(* IEC 61131-3 sources: daoli-st-library/DL_Algo (part 18) *)

(* ---- FB_DL_PidController.st ---- *)
(*==============================================================================
 * 组件名称 (Component)  : FB_DL_PidController
 * 所属子库 (Sublibrary) : DL_Algo
 * 当前版本 (Version)    : 1.0.1
 * 兼容性   (Platform)   : CODESYS 3.5 / TwinCAT 3 / 汇川 InoProShop / Machine Expert
 *                         仅依赖 Standard.library（R_TRIG），零厂商方言
 * 功能描述 (Function)   : 单回路通用离散 PID 控制器。位置式与增量式由独立布尔
 *                         bIncremental 选择（不堆模式枚举）；含控制死区、积分
 *                         分离（触限停积分）、两级抗积分饱和（条件积分 + 限幅
 *                         反算回填）、手自动无扰切换与跟踪回投。fKp 为负即反
 *                         作用（沿 OSCAT / 西门子惯例）。现场用途：温度 / 压力 /
 *                         流量单闭环调节主块，温控区与后续串级块的基石。
 * 开源溯源 (Origin)     : 原创实现。功能分类与参数域参考 OSCAT 基础库 FT_PIWL
 *                         反算抗饱和思想与西门子 CONT_C 公开语义描述，
 *                         未复制任何厂商源码，clean-room 重写。
 * 本文件内含       : TYPE  E_DL_PidState（配套枚举，归属 DL_Algo）
 *                    FB    FB_DL_PidController
 * 依赖     (Depends)    : 无 DL_ 内部依赖；Standard.library: R_TRIG
 * 红线自检 (Redline)    : R1 ✓ 零全局变量表与外部变量引用 ｜ R2 ✓ 零物理 IO 地址直写
 *                         R3 ✓ 纯 IEC 61131-3 ｜ R4 ✓ 防除零+钳位+非有限值防御
 *                         R5 ✓ 全变量中英双语同行注释 ｜ R6 ✓ 四态 ENUM+CASE+ELSE
 *                         R7 ✓ R_TRIG 实例主体最前部无条件刷新
 * 修订历史 (Revision)   :
 *   2026-11-15  v1.0.0  首版入库 · Round 04 · Level 1 DL_Algo
 *   2026-11-15  v1.0.1  阶段五终审精修：积分量纲统一为[%]；eIdle 补 bActive
 *                       清零；信息级码不置 bError；首扫与手自动历史同步防踢腿
 * 验收向量 (Acceptance) :
 *   V1 阶跃纯比例：fKp=2, tTi=T#0S, SP=50, PV=0 → fOut=rOutMax 触限
 *   V2 抗饱和：fKp=2, tTi=T#2S, SP=200 → 触上限后撤销阶跃，输出快速回落
 *      （积分已反算回填，无长时间停限）
 *   V3 无扰切换：手动 30.0 切自动首拍输出保持 30.0 连续
 *   V4 死区：fDeadband=5 且 |偏差|<5 → 输出保持不变
 *   V5 非有限值：fSetpoint 写入非法浮点 → 输出保持上一拍且 uErrorId=0002_0004
 *   V6 增量式：fKp=1, tTi=T#1S, 恒偏差 10 → fOut 单调爬升至上限后停
 *============================================================================*)
(*-----------------------------------------------------------------------------
 * 枚举: E_DL_PidState（归属 DL_Algo，与 FB_DL_PidController 同文件）
 * 含义: PID 控制器离散状态。数值步长留空位便于后续插态而不破坏已有工程。
 *----------------------------------------------------------------------------*)
TYPE E_DL_PidState :
(
    eIdle   := 0,    // 使能关：输出回输出下限，积分冻结 / Idle: enable off, output at low limit, integral frozen
    eAuto   := 10,   // 自动调节：闭环 PID 运算中 / Auto: closed-loop PID computation active
    eManual := 20,   // 手动模式：输出手动值，积分同步跟踪保证无扰 / Manual: output manual value, integral tracked for bumpless
    eFault  := 99    // 故障兜底态：非法状态进入，输出安全值 / Fault fallback: entered on illegal state, safe output
);
END_TYPE
(*==============================================================================
 * 功能块: FB_DL_PidController
 * 调用约定: 每个扫描周期无条件调用一次；bReset 上升沿清积分与故障。
 * 无状态泄漏: 全部状态驻留于实例私有 VAR，零全局引用，可多实例并行。
 * 工程披露: 微分项对偏差做一阶预滤波（滤波时间取 tTd 的 1/10），抑制微分尖峰。
 *============================================================================*)
FUNCTION_BLOCK FB_DL_PidController
VAR_INPUT
    bEnable      : BOOL := FALSE;     // 总使能，FALSE 时输出回输出下限 / Master enable, FALSE drives output to low limit
    bManual      : BOOL := FALSE;     // 手动模式选择，TRUE = 手动输出 / Manual mode select, TRUE = manual output
    fManualValue : REAL := 0.0;       // 手动输出值 [%]，越限自动钳位 / Manual output value [%], auto-clamped
    fSetpoint    : REAL := 0.0;       // 设定值 [EU] / Setpoint in engineering units
    fActual      : REAL := 0.0;       // 过程实际值 [EU] / Process actual value in engineering units
    fKp          : REAL := 1.0;       // 比例增益 [1]，负值 = 反作用 / Proportional gain, negative = reverse acting
    tTi          : TIME := T#2S;      // 积分时间 [s]，T#0S 表示纯 PD 无积分 / Integral time [s], T#0S = pure PD
    tTd          : TIME := T#0S;      // 微分时间 [s]，T#0S 关闭微分 / Derivative time [s], T#0S disables derivative
    fDeadband    : REAL := 0.0;       // 控制死区 [EU]，负值自动钳 0 / Control deadband [EU], negative clamped to 0
    bIncremental : BOOL := FALSE;     // TRUE = 增量式算法，FALSE = 位置式 / TRUE = incremental form, FALSE = positional
    rOutMin      : REAL := 0.0;       // 输出下限 [%] / Output lower limit in percent
    rOutMax      : REAL := 100.0;     // 输出上限 [%] / Output upper limit in percent
    tSampleTime  : TIME := T#100MS;   // 采样周期 [s]，小于 T#10MS 钳位 / Sample period, clamped to 10 ms minimum
    bTrack       : BOOL := FALSE;     // 跟踪使能，TRUE 时输出立即跟随跟踪值 / Track enable, output follows track value
    fTrackValue  : REAL := 0.0;       // 跟踪值 [%]，与输出同量纲，用于无扰投切 / Track value in percent, same unit as output
    bReset       : BOOL := FALSE;     // 复位信号，上升沿清积分与故障 / Reset, rising edge clears integral and fault
END_VAR
VAR_OUTPUT
    fOut         : REAL;              // 控制输出 [%] / Control output in percent
    fErr         : REAL;              // 偏差 = 设定 - 实际 [EU] / Error = setpoint minus actual
    fIntPart     : REAL;              // 积分分量 [%]，诊断用 / Integral component in percent, diagnostics
    bLimitHigh   : BOOL;              // 输出触上限标志 / Output saturated at upper limit flag
    bLimitLow    : BOOL;              // 输出触下限标志 / Output saturated at lower limit flag
    bActive      : BOOL;              // 自动调节进行中标志 / Auto regulation active flag
    bError       : BOOL;              // 故障标志，0 除外均置位 / Fault flag, set on any nonzero error code
    uErrorId     : UDINT;             // 故障码，0 = 无故障 / Error code, 0 = no error
END_VAR
VAR
    fErrPrev1    : REAL;              // 上一拍偏差（增量式历史） [EU] / Previous error for incremental form
    fErrPrev2    : REAL;              // 上上拍偏差（增量式历史） [EU] / Error two cycles ago for incremental form
    fErrF        : REAL;              // 微分预滤波后的偏差 [EU] / Prefiltered error for derivative term
    fErrFPrev    : REAL;              // 上一拍预滤波偏差 [EU] / Previous prefiltered error
    fbTrigReset  : R_TRIG;            // 复位信号上升沿检测实例 / Reset rising edge detector instance
    eState       : E_DL_PidState;     // 主状态机当前状态 / Current state of the main state machine
    bInit        : BOOL := TRUE;      // 历史同步标志，TRUE 触发历史同步（首扫即同步防踢腿）/ History sync flag, TRUE syncs histories on first scan
    fDt          : REAL;              // 生效采样周期 [s] / Effective sample period in seconds
    fLimLow      : REAL;              // 修复后的输出下限 [%] / Repaired output lower limit
    fLimHigh     : REAL;              // 修复后的输出上限 [%] / Repaired output upper limit
    fDeadbandEff : REAL;              // 钳位后的有效死区 [EU] / Clamped effective deadband
    fInt         : REAL;              // 积分累积 [%]，与输出同量纲 / Accumulated integral in percent, same unit as output
    fP           : REAL;              // 比例分量 [%] / Proportional component
    fD           : REAL;              // 微分分量 [%] / Derivative component
    fPre         : REAL;              // 抗饱和判定用预输出 [%] / Pre-output for anti-windup test
    fDelta       : REAL;              // 增量式单拍增量 [%] / Incremental delta of one cycle
    fTdS         : REAL;              // 微分时间换算秒 [s] / Derivative time in seconds
    fAlpha       : REAL;              // 微分预滤波权重 [0..1] / Derivative prefilter weight
    fManOut      : REAL;              // 钳位后的手动输出 [%] / Clamped manual output
    bSkipInt     : BOOL;              // 积分分离标志：触限且误差继续推进 / Conditional integration flag
END_VAR
VAR CONSTANT
    DL_PID_ERR_MAX : REAL := 1.0E10;  // 积分钳位上限 [%]，防浮点溢出的极端钳位 / Integral clamp ceiling [%], extreme guard against float overflow
END_VAR
(*------------------------------------------------------------------------------
 * 段 1｜无条件刷新区（红线 R7）：复位沿检测严禁进入任何 IF / CASE 分支
 *      Unconditional refresh zone (red line R7): edge detector outside IF / CASE
 *-----------------------------------------------------------------------------*)
fbTrigReset(CLK := bReset);
(*------------------------------------------------------------------------------
 * 段 2｜参数钳位与公共防御（不中断扫描，现场组态笔误不停机）
 *      Parameter clamping and common defenses, never stops the scan
 *-----------------------------------------------------------------------------*)
bError   := FALSE;                    // 每拍重算故障标志 / Recompute fault flag every cycle
uErrorId := 16#0002_0000;             // 每拍重算故障码 / Recompute error code every cycle
bLimitHigh := FALSE;                  // 触限标志每拍重算 / Saturation flags recomputed every cycle
bLimitLow  := FALSE;                  // 触限标志每拍重算 / Saturation flags recomputed every cycle
IF tSampleTime < T#10MS THEN
    fDt := 0.01;                      // 采样周期非法钳位为 0.01 s / Illegal sample period clamped to 0.01 s
    uErrorId := 16#0002_0002;         // 公共码：采样周期已钳位 / Common code: sample period clamped
ELSE
    fDt := TIME_TO_REAL(tSampleTime) / 1000.0;  // 采样周期换算为秒 [s] / Sample period converted to seconds
END_IF
IF rOutMin > rOutMax THEN
    fLimLow  := rOutMax;              // 上下限对调修复（下限取原上限） / Swapped limits after repair
    fLimHigh := rOutMin;              // 上下限对调修复（上限取原下限） / Swapped limits after repair
    uErrorId := 16#0002_0001;         // 公共码：参数越界已钳位 / Common code: parameter clamped
ELSE
    fLimLow  := rOutMin;              // 合法下限直通 / Valid lower limit passed through
    fLimHigh := rOutMax;              // 合法上限直通 / Valid upper limit passed through
END_IF
IF fDeadband < 0.0 THEN
    fDeadbandEff := 0.0;              // 死区负值钳 0 / Negative deadband clamped to zero
    uErrorId := 16#0002_0001;         // 公共码：参数越界已钳位 / Common code: parameter clamped
ELSE
    fDeadbandEff := fDeadband;        // 合法死区直通 / Valid deadband passed through
END_IF
(*------------------------------------------------------------------------------
 * 段 3｜复位处理：清积分、清增量式历史、清滤波偏差，故障归零
 *      Reset handling: clear integral, incremental history and filtered error
 *-----------------------------------------------------------------------------*)
IF fbTrigReset.Q THEN
    fInt       := 0.0;                // 清积分累积 [%] / Clear accumulated integral in percent
    fErrPrev1  := 0.0;                // 清上一拍偏差 / Clear previous error history
    fErrPrev2  := 0.0;                // 清上上拍偏差 / Clear two-cycle error history
    fErrF      := 0.0;                // 清滤波偏差 / Clear prefiltered error
    fErrFPrev  := 0.0;                // 清上拍滤波偏差 / Clear previous prefiltered error
    fOut       := fLimLow;            // 输出回安全下限 / Output to safe lower limit
    eState     := eIdle;              // 状态回空闲 / State back to idle
    bInit      := TRUE;               // 置首扫标志使下一拍同步历史 / Set init flag to resync history next cycle
END_IF
(*------------------------------------------------------------------------------
 * 段 4｜非有限值防御：设定值 / 过程值 / 手动值 / 跟踪值任一非法即拒绝本拍更新
 *      Non-finite defense: reject this cycle if any relevant input is invalid
 *-----------------------------------------------------------------------------*)
IF (fSetpoint <> fSetpoint) OR (ABS(fSetpoint) > 1.0E30)
   OR (fActual <> fActual) OR (ABS(fActual) > 1.0E30)
   OR (fManualValue <> fManualValue) OR (ABS(fManualValue) > 1.0E30)
   OR (fTrackValue <> fTrackValue) OR (ABS(fTrackValue) > 1.0E30) THEN
    bError   := TRUE;                 // 置故障标志 / Set fault flag
    uErrorId := 16#0002_0004;         // 公共码：输入非有限值已拒绝 / Common code: non-finite input rejected
    RETURN;                           // 保持上一拍输出与状态 / Hold previous output and state
END_IF
(*------------------------------------------------------------------------------
 * 段 5｜使能关断：输出回下限、积分冻结、状态回空闲（允许带电观察）
 *      Enable off: output to low limit, integral frozen, state back to idle
 *-----------------------------------------------------------------------------*)
IF NOT bEnable THEN
    eState  := eIdle;                 // 强制回空闲态 / Force idle state
    fOut    := fLimLow;               // 输出回下限安全值 / Output to safe low limit
    fErr    := fSetpoint - fActual;   // 偏差仍刷新供诊断 / Error still refreshed for diagnostics
    bActive := FALSE;                 // 调节未激活 / Regulation not active
    fIntPart:= fInt;                  // 保留积分分量供诊断 / Keep integral component for diagnostics
    RETURN;                           // 本拍结束 / End of this cycle
END_IF
(*------------------------------------------------------------------------------
 * 段 6｜主状态机（红线 R6）：ENUM + CASE + ELSE 兜底
 *      Main state machine: ENUM + CASE with mandatory ELSE fallback
 *-----------------------------------------------------------------------------*)
CASE eState OF
    eIdle:
        (* 空闲态：按手动 / 自动请求迁移，迁移前同步增量式历史防微分踢腿 *)
        (* Idle: migrate by mode request, sync incremental history before transfer *)
        bActive := FALSE;             // 空闲态激活标志清零防跨拍残留 / Clear active flag against stale carry-over
        fErr := fSetpoint - fActual;  // 计算原始偏差 [EU] / Raw error in engineering units
        IF ABS(fErr) < fDeadbandEff THEN
            fErr := 0.0;              // 死区内偏差按 0 处理 / Error inside deadband treated as zero
        END_IF
        IF bManual THEN
            eState := eManual;        // 请求手动 / Request manual mode
        ELSE
            eState := eAuto;          // 请求自动 / Request auto mode
        END_IF
    eAuto:
        (* 自动调节态：位置式或增量式 PID 闭环运算 + 两级抗饱和 *)
        (* Auto: positional or incremental closed-loop PID with two-stage anti-windup *)
        bActive := TRUE;              // 自动调节激活 / Auto regulation active
        fErr := fSetpoint - fActual;  // 原始偏差 [EU] / Raw error
        IF ABS(fErr) < fDeadbandEff THEN
            fErr := 0.0;              // 死区内偏差置 0 / Zero error inside deadband
        END_IF
        IF bInit THEN
            (* 首扫 / 复位后同步全部历史，杜绝上电尖峰与虚假微分 *)
            (* First scan / post-reset history sync, no power-up spike *)
            fErrF     := fErr;        // 滤波偏差同步 / Sync prefiltered error
            fErrFPrev := fErr;        // 上拍滤波偏差同步 / Sync previous prefiltered error
            fErrPrev1 := fErr;        // 增量式历史同步 / Sync incremental history
            fErrPrev2 := fErr;        // 增量式历史同步 / Sync incremental history
            bInit     := FALSE;       // 清首扫标志 / Clear first-scan flag
        END_IF
        fP := fKp * fErr;             // 比例项 [%] / Proportional term
        IF bTrack THEN
            (* 跟踪回投：输出立即跟随跟踪值，积分反算同步，恢复自动零扰动 *)
            (* Track mode: output follows track value, integral back-calculated in sync *)
            fOut    := LIMIT(fLimLow, fTrackValue, fLimHigh);   // 输出钳位跟随 / Clamped tracking output
            fInt    := fOut - fP - fD;                          // 积分反算同步 / Back-calculated integral
            fErrF   := fErr;        // 滤波偏差同步 / Sync prefiltered error
            fErrFPrev := fErr;      // 上拍滤波偏差同步 / Sync previous prefiltered error
            fErrPrev1 := fErr;      // 增量式历史同步 / Sync incremental history
            fErrPrev2 := fErr;      // 增量式历史同步 / Sync incremental history
            fIntPart := fInt;       // 诊断分量刷新 / Refresh diagnostic component
        ELSIF bIncremental THEN
            (* 增量式：PID 增量作用于输出累积，天然抗饱和由限幅兜底 *)
            (* Incremental form: PID delta applied to output accumulation *)
            fDelta := fKp * (fErr - fErrPrev1);                 // 比例增量 [%] / Proportional delta
            IF tTi > T#0S THEN
                fDelta := fDelta + fKp * fErr * fDt / (TIME_TO_REAL(tTi) / 1000.0);  // 积分增量 / Integral delta
            END_IF
            IF tTd > T#0S THEN
                fDelta := fDelta + fKp * (TIME_TO_REAL(tTd) / 1000.0) / fDt
                          * (fErr - 2.0 * fErrPrev1 + fErrPrev2);  // 微分增量 / Derivative delta
            END_IF
            fOut := LIMIT(fLimLow, fOut + fDelta, fLimHigh);    // 输出累积并限幅 / Accumulate and clamp
            fErrPrev2 := fErrPrev1;                             // 历史滚动 / Roll history
            fErrPrev1 := fErr;                                  // 历史滚动 / Roll history
            fIntPart  := fOut - fP - fD;                        // 诊断分量 / Diagnostic component
            IF ((fOut >= fLimHigh) AND (fDelta > 0.0))
               OR ((fOut <= fLimLow) AND (fDelta < 0.0)) THEN
                bLimitHigh := (fOut >= fLimHigh);               // 触上限标志 / Upper saturation flag
                bLimitLow  := (fOut <= fLimLow);                // 触下限标志 / Lower saturation flag
                IF uErrorId = 16#0002_0000 THEN
                    uErrorId := 16#0002_0101;                   // 信息级：输出饱和提示 / Info: output saturated
                END_IF
            END_IF
        ELSE
            (* 位置式：先做微分预滤波，再做积分分离与两级抗饱和 *)
            (* Positional: derivative prefilter, then conditional integration and back-calc *)
            IF tTd > T#0S THEN
                fTdS   := TIME_TO_REAL(tTd) / 1000.0;           // 微分时间换算秒 [s] / Derivative time in seconds
                fAlpha := fDt / (0.1 * fTdS + fDt);             // 预滤波权重 [0..1] / Prefilter weight
                fErrF  := fErrF + fAlpha * (fErr - fErrF);      // 一阶预滤波递推 / First-order prefilter recursion
                fD     := fKp * fTdS / fDt * (fErrF - fErrFPrev);  // 微分项 [%] / Derivative term
                fErrFPrev := fErrF;                             // 滚动滤波历史 / Roll filtered history
            ELSE
                fD        := 0.0;                               // 微分关闭 / Derivative disabled
                fErrF     := fErr;                              // 滤波偏差直通 / Prefiltered error follows
                fErrFPrev := fErr;                              // 上拍滤波偏差同步 / Sync previous value
            END_IF
            fPre := fP + fD + fInt;                             // 当前积分下的预输出 [%] / Pre-output with current integral
            bSkipInt := (fPre > fLimHigh AND fErr > 0.0)
                     OR (fPre < fLimLow  AND fErr < 0.0);       // 积分分离判定 / Conditional integration test
            IF (tTi > T#0S) AND (NOT bSkipInt) THEN
                fInt := fInt + fKp * fErr * fDt / (TIME_TO_REAL(tTi) / 1000.0);  // 条件积分 / Conditional integration
            END_IF
            fInt := LIMIT(-DL_PID_ERR_MAX, fInt, DL_PID_ERR_MAX);  // 积分钳位防溢出 / Clamp integral against overflow
            fPre := fP + fD + fInt;                             // 二次合成预输出 [%] / Recomposed pre-output
            IF fPre > fLimHigh THEN
                fOut := fLimHigh;                               // 输出钳上限 / Output at upper limit
                fInt := fLimHigh - fP - fD;                     // 反算回填积分 / Back-calculated integral
                bLimitHigh := TRUE;                             // 触上限标志 / Upper saturation flag
                IF uErrorId = 16#0002_0000 THEN
                    uErrorId := 16#0002_0101;                   // 信息级：输出饱和提示 / Info: output saturated
                END_IF
            ELSIF fPre < fLimLow THEN
                fOut := fLimLow;                                // 输出钳下限 / Output at lower limit
                fInt := fLimLow - fP - fD;                      // 反算回填积分 / Back-calculated integral
                bLimitLow := TRUE;                              // 触下限标志 / Lower saturation flag
                IF uErrorId = 16#0002_0000 THEN
                    uErrorId := 16#0002_0101;                   // 信息级：输出饱和提示 / Info: output saturated
                END_IF
            ELSE
                fOut := fPre;                                   // 正常输出 / Normal output
            END_IF
            fIntPart := fInt;                                   // 诊断分量刷新 / Refresh diagnostic component
        END_IF
        IF bManual THEN
            eState := eManual;                                  // 切手动 / Switch to manual
        END_IF
    eManual:
        (* 手动态：输出手动值（钳位），积分反算同步保证回自动瞬间输出连续 *)
        (* Manual: clamped manual output, integral back-calculated for bumpless return *)
        bActive := FALSE;                                       // 自动调节未激活 / Auto not active
        fErr := fSetpoint - fActual;                            // 偏差仍计算供诊断 / Error for diagnostics
        IF ABS(fErr) < fDeadbandEff THEN
            fErr := 0.0;                                        // 死区内偏差置 0 / Zero inside deadband
        END_IF
        (* 手动期间持续同步微分与增量式历史，杜绝切回自动瞬间的踢腿 *)
        (* Keep syncing derivative and incremental history in manual, no kick on auto return *)
        fErrF     := fErr;                                      // 微分滤波偏差同步 / Sync prefiltered error
        fErrFPrev := fErr;                                      // 上拍滤波偏差同步 / Sync previous prefiltered error
        fErrPrev1 := fErr;                                      // 增量式历史同步 / Sync incremental history
        fErrPrev2 := fErr;                                      // 增量式历史同步 / Sync incremental history
        fP := fKp * fErr;                                       // 比例项 [%] / Proportional term
        fD := 0.0;                                              // 手动下微分置 0 / Derivative zero in manual
        fManOut := LIMIT(fLimLow, fManualValue, fLimHigh);      // 手动值钳位 / Clamped manual value
        IF fManualValue > fLimHigh OR fManualValue < fLimLow THEN
            IF uErrorId = 16#0002_0000 THEN
                uErrorId := 16#0002_0102;                       // 手动值超限已钳位 / Manual value clamped
            END_IF
        END_IF
        fOut      := fManOut;                                   // 输出手动值 / Output manual value
        fInt      := fManOut - fP - fD;                         // 积分反算同步 / Back-calculated integral
        fInt      := LIMIT(-DL_PID_ERR_MAX, fInt, DL_PID_ERR_MAX);  // 积分钳位 / Clamp integral
        fIntPart  := fInt;                                      // 诊断分量刷新 / Refresh diagnostic component
        IF bTrack THEN
            fOut := LIMIT(fLimLow, fTrackValue, fLimHigh);      // 跟踪值优先 / Track value takes priority
            fInt := fOut - fP - fD;                             // 积分同步 / Integral in sync
        END_IF
        IF bInit THEN
            fErrF     := fErr;                                  // 滤波偏差同步 / Sync prefiltered error
            fErrFPrev := fErr;                                  // 上拍滤波偏差同步 / Sync previous value
            fErrPrev1 := fErr;                                  // 增量式历史同步 / Sync history
            fErrPrev2 := fErr;                                  // 增量式历史同步 / Sync history
            bInit     := FALSE;                                 // 清首扫标志 / Clear first-scan flag
        END_IF
        IF NOT bManual THEN
            eState := eAuto;                                    // 切自动 / Switch to auto
        END_IF
    eFault:
        (* 故障兜底态：输出安全下限，等待复位沿解除 *)
        (* Fault fallback: safe low-limit output, released by reset edge *)
        fOut    := fLimLow;                                     // 安全输出 / Safe output
        bActive := FALSE;                                       // 调节未激活 / Not active
    ELSE
        (* 非法状态拦截：任何未定义状态一律进故障兜底，不做隐式恢复 *)
        (* Illegal state interception: any undefined state goes to fault fallback *)
        eState   := eFault;                                     // 进故障态 / Enter fault state
        bError   := TRUE;                                       // 置故障标志 / Set fault flag
        uErrorId := 16#0002_0005;                               // 非法状态兜底码 / Illegal state fallback code
        fOut     := fLimLow;                                    // 安全输出 / Safe output
END_CASE;
(* 信息级码（0101 输出饱和 / 0102 手动值钳位）不置故障标志，防下游报警误动作 *)
(* Info-level codes (saturation / manual clamp) never raise the fault flag *)
bError := (uErrorId <> 16#0002_0000) AND (uErrorId <> 16#0002_0101)
          AND (uErrorId <> 16#0002_0102);                        // 非信息级码才置故障 / Fault flag only on non-info codes
END_FUNCTION_BLOCK

(* ---- FB_DL_PidGainScheduler.st ---- *)
(*==============================================================================
 * 组件名称 (Component)  : FB_DL_PidGainScheduler
 * 溯源说明 (Provenance) : 道莅 clean-room 防御性实现（LGF Technology 深化 + 规划新增线）
 * 所属子库 (Sublibrary) : DL_Algo / ControlParams
 * 当前版本 (Version)    : 1.0.0
 * 兼容性   (Platform)   : CODESYS 3.5 / TwinCAT 3 / 汇川 InoProShop；
 *                         纯 IEC 61131-3（第 3 版），零标准库依赖
 * 组件分类 (Category)   : 功能块（FUNCTION_BLOCK）· 增益调度查表插值
 * 功能一句话 (Summary)  : 按调度变量查增益表线性插值输出 Kp/Ti/Td，仅出参数不控回路。
 * 边界与安全 (Boundary) : ①调度变量低于首点/高于末点 → 端点钳位并置码 3705；
 *                         ②表未按 fVar 严格升序 → 码 3701 且 bHoldLast 生效保持上次输出；
 *                         ③调度变量 NaN → 码 3702 保持上次输出；
 *                         ④表点数不足 2 → 视同表非法（3701 复用）；
 *                         ⑤本件只产出参数，不内嵌控制回路（与 PID 件正交解耦）。
 * 错误码    : 16#0002_3701 增益表非法（未升序或点数不足）——故障级（持续态）
 *             16#0002_3702 调度变量 NaN（保持上次输出）——故障级（持续态）
 *             16#0002_3705 端点钳位发生——信息级（持续态）
 * 码位总账  : 16#0002_3701 用 / 16#0002_3702 用 / 16#0002_3705 用
 * 修改记录  : v1.0.0 R26 初版
 *==============================================================================*)
TYPE ST_DL_GainPoint :
STRUCT
    fVar : LREAL; // 调度变量锚点 / Scheduling variable anchor
    fKp  : LREAL; // 该锚点比例增益 / Proportional gain at anchor
    fTi  : LREAL; // 该锚点积分时间 [s] / Integral time at anchor [s]
    fTd  : LREAL; // 该锚点微分时间 [s] / Derivative time at anchor [s]
END_STRUCT
END_TYPE

FUNCTION_BLOCK FB_DL_PidGainScheduler
VAR_INPUT
    fSchedVar  : LREAL; // 调度变量（如流量/温度工况）/ Scheduling variable
    bEnable    : BOOL;  // 使能：FALSE 保持上次输出 / Enable: FALSE holds last output
    bHoldLast  : BOOL;  // 表非法时保持上次输出 / Hold last output on illegal table
END_VAR
VAR_IN_OUT
    aGainTable : ARRAY[*] OF ST_DL_GainPoint; // 增益表，须按 fVar 升序 / Gain table, ascending by fVar
END_VAR
VAR_OUTPUT
    fKp   : LREAL; // 插值输出比例增益 / Interpolated proportional gain
    fTi   : LREAL; // 插值输出积分时间 [s] / Interpolated integral time [s]
    fTd   : LREAL; // 插值输出微分时间 [s] / Interpolated derivative time [s]
    eErr  : UDINT; // 本周期错误码，0=无错 / Error code this cycle, 0 = none
END_VAR
VAR
    nPts    : INT;  // 表点数 / Table point count
    i       : INT;  // 分段搜索游标 / Segment search cursor
    fDen    : LREAL; // 分段分母（前判零）/ Segment denominator (zero-guarded)
    fRatio  : LREAL; // 段内插值比例 / Interpolation ratio
    bTableOk: BOOL; // 表合法性中间判据 / Table legality intermediate
    bHold   : BOOL; // 本拍保持输出判据 / Hold-output predicate this cycle
END_VAR

// ---------- 周期起点：错误码清零（持续态随后重置） ----------
eErr := 0;
bHold := FALSE;

// ---------- 使能为假：纯保持，不查表不刷新 ----------
IF NOT bEnable THEN
    bHold := TRUE;                            // 保持上次输出 / Hold last output
ELSE
    // ---------- 表点数与单调性防御 ----------
    nPts := UPPER_BOUND(aGainTable, 1) + 1;   // 表点数 / Point count
    bTableOk := nPts >= 2;                    // 至少两点 / At least two points
    IF bTableOk THEN
        FOR i := 0 TO nPts - 2 DO
            IF NOT (aGainTable[i].fVar < aGainTable[i + 1].fVar) THEN
                bTableOk := FALSE;            // 严格升序被破坏 / Strict order violated
            END_IF
        END_FOR
    END_IF
    IF NOT bTableOk THEN
        eErr  := 16#0002_3701;                // 表非法码 / Illegal table code
        bHold := bHoldLast;                   // 按调用方策略保持 / Hold per caller policy
    ELSE
        // ---------- NaN 调度变量：保持 ----------
        IF fSchedVar <> fSchedVar THEN
            eErr  := 16#0002_3702;            // NaN 码 / NaN code
            bHold := TRUE;                    // 强制保持 / Forced hold
        ELSE
            // ---------- 端点钳位与段内插值 ----------
            IF fSchedVar <= aGainTable[0].fVar THEN
                fKp := aGainTable[0].fKp;     // 低于首点钳端点 / Below first: clamp endpoint
                fTi := aGainTable[0].fTi;
                fTd := aGainTable[0].fTd;
                IF fSchedVar < aGainTable[0].fVar THEN
                    eErr := 16#0002_3705;     // 端点钳位码 / Endpoint clamp code
                END_IF
            ELSIF fSchedVar >= aGainTable[nPts - 1].fVar THEN
                fKp := aGainTable[nPts - 1].fKp; // 高于末点钳端点 / Above last: clamp endpoint
                fTi := aGainTable[nPts - 1].fTi;
                fTd := aGainTable[nPts - 1].fTd;
                IF fSchedVar > aGainTable[nPts - 1].fVar THEN
                    eErr := 16#0002_3705;     // 端点钳位码 / Endpoint clamp code
                END_IF
            ELSE
                i := 0;
                WHILE (i < nPts - 2) AND (fSchedVar > aGainTable[i + 1].fVar) DO
                    i := i + 1;               // 定位所在段 / Locate segment
                END_WHILE
                fDen := aGainTable[i + 1].fVar - aGainTable[i].fVar; // 段宽 / Segment width
                IF fDen > 0.0 THEN
                    fRatio := (fSchedVar - aGainTable[i].fVar) / fDen; // 除法前判零 / Zero-guarded divide
                    fKp := aGainTable[i].fKp + fRatio * (aGainTable[i + 1].fKp - aGainTable[i].fKp);
                    fTi := aGainTable[i].fTi + fRatio * (aGainTable[i + 1].fTi - aGainTable[i].fTi);
                    fTd := aGainTable[i].fTd + fRatio * (aGainTable[i + 1].fTd - aGainTable[i].fTd);
                ELSE
                    fKp := aGainTable[i].fKp; // 段宽为零防御取左点 / Zero-width defensive left point
                    fTi := aGainTable[i].fTi;
                    fTd := aGainTable[i].fTd;
                END_IF
            END_IF
        END_IF
    END_IF
END_IF

// ---------- 保持路径显式化：bHold 时三输出不动（锁存语义注释） ----------
// bHold=TRUE 期间 fKp/fTi/fTd 为上次有效锁存值，内部不引入实时镜像副本，
// 输出与内部判定共用同一组锁存变量，避免双口径混用。

END_FUNCTION_BLOCK

(* ---- FB_DL_PidParamDriftAudit.st ---- *)
(*
  Name        : FB_DL_PidParamDriftAudit
  Category    : DL_Algo
  Version     : 1.0.1
  Purpose     : 整定参数漂移审计：逐拍比对现行 Kp/Ti/Td 与基准快照，按相对容差判漂移并累计越差次数，供「谁改了参数」留痕；/ Audit PID parameter drift: compare live Kp/Ti/Td against baseline snapshots with relative tolerance, accumulate excursions for an auditable trail
  溯源        : 借 t2-3-风格指南·审计 的分类/参数域组织，clean-room 实现
  Boundary    : ① 基准近零分支：|基准| <= eps 时相对偏差无定义，改走绝对差判据（fTolAbs），不产生除零/Inf；
                ② 现行与基准同为近零 → 判无漂移（0/0 语义按「一致」处理）；
                ③ 容差与近零判据全部 ABS 差比较，禁 `=`/`<>`；
                ④ 越差计数饱和累加，防 UDINT 回绕；
                ⑤ 本件只审计不改参数，输出仅供上位留痕（属主边界）。
  修订记录    : 2026-11-20 v1.0.1：六参数有限性闸补 Inf 差判（NaN+Inf 双闸，R52-05）；bDriftAny 改由三确认位 OR 同源重算（R52-06）；_fHun 迁入 VAR CONSTANT c_fHun 收口魔法数。
*)
TYPE E_DL_PdaState :
(
    eIdle  := 0,                             (* 未使能 / Disabled *)
    eAudit := 10,                            (* 审计运行 / Auditing *)
    eFault := 90                             (* 故障锁存相 / Fault latched *)
);
END_TYPE

TYPE E_DL_PdaCause :
(
    eNone       := 0,                        (* 无故障成因 / No cause *)
    eCfgIllegal := 1,                        (* 组态非法：容差/参考值越域 / Illegal config *)
    ePhaseBad   := 2                         (* 非法相位兜底 / Illegal phase fallback *)
);
END_TYPE

FUNCTION_BLOCK FB_DL_PidParamDriftAudit
VAR_INPUT
    fKp        : REAL := 1.0;                (* 现行比例增益 [-] / Live proportional gain *)
    fTi        : REAL := 1.0;                (* 现行积分时间，P 模式可为 0 [s] / Live integral time, 0 allowed *)
    fTd        : REAL := 0.0;                (* 现行微分时间，P/PI 模式可为 0 [s] / Live derivative time, 0 allowed *)
    fKpRef     : REAL := 1.0;                (* 基准比例增益（签核快照）[-] / Baseline proportional gain *)
    fTiRef     : REAL := 1.0;                (* 基准积分时间 [s] / Baseline integral time *)
    fTdRef     : REAL := 0.0;                (* 基准微分时间 [s] / Baseline derivative time *)
    fTolRel    : REAL := 0.05;               (* 相对漂移容差（5% = 0.05），域 > 0 [-] / Relative tolerance, > 0 *)
    fTolAbs    : REAL := 0.01;               (* 基准近零时改用的绝对差容差，域 > 0 [参数单位] / Absolute tolerance for near-zero baselines *)
    nConfirm   : INT := 3;                   (* 越差确认拍数，域 >= 1 [拍] / Consecutive excursion scans to confirm *)
    bEnable    : BOOL := TRUE;               (* 审计使能 [-] / Enable *)
    bReset      : BOOL := FALSE;             (* 复位命令，上升沿清漂移标志与计数 [-] / Reset command *)
END_VAR
VAR_OUTPUT
    fDriftKp   : REAL;                       (* Kp 相对漂移（% / 近零基准时为绝对差）[%] / Kp drift *)
    fDriftTi   : REAL;                       (* Ti 相对漂移 [%] / Ti drift *)
    fDriftTd   : REAL;                       (* Td 相对漂移 [%] / Td drift *)
    bDriftKp   : BOOL;                       (* Kp 越差确认位 [-] / Kp drift confirmed *)
    bDriftTi   : BOOL;                       (* Ti 越差确认位 [-] / Ti drift confirmed *)
    bDriftTd   : BOOL;                       (* Td 越差确认位 [-] / Td drift confirmed *)
    bDriftAny  : BOOL;                       (* 任一参数越差（汇总位）[-] / Any parameter drifted *)
    nDriftCnt  : UDINT;                      (* 累计确认越差次数（饱和）[-] / Confirmed drift count, saturated *)
    eState     : E_DL_PdaState;              (* 状态出口 / State outlet *)
    eCause     : E_DL_PdaCause;              (* 故障成因出口（R190 归因唯一） / Fault cause outlet *)
    bError     : BOOL;                       (* 故障锁存标志 [-] / Fault latch flag *)
END_VAR
VAR
    _eState  : E_DL_PdaState := E_DL_PdaState.eIdle;     (* 内部相位（CASE 唯一写入目标） / Internal phase *)
    _eCause  : E_DL_PdaCause := E_DL_PdaCause.eNone;     (* 故障成因锁存量 / Latched cause *)
    rtReset  : R_TRIG;                       (* 复位沿实例，段 0 无条件调用 / Reset edge instance *)
    _bFault  : BOOL;                         (* 故障锁存位 / Latched fault bit *)
    _bCfgBad : BOOL;                         (* 组态非法当拍量 / Illegal config this scan *)
    _bFinite : BOOL;                         (* 六参数有限性联合闸 / Finiteness of all six parameters *)
    _bExKp   : BOOL;                         (* Kp 当拍越差（未确认） / Kp excursion this scan *)
    _bExTi   : BOOL;                         (* Ti 当拍越差 / Ti excursion this scan *)
    _bExTd   : BOOL;                         (* Td 当拍越差 / Td excursion this scan *)
    _bAny    : BOOL;                         (* 任一当拍越差 / Any excursion this scan *)
    _nHold   : INT;                          (* 越差连续拍计数 [-] / Consecutive excursion counter *)
    _fDkp    : REAL;                         (* Kp 偏差绝对值/相对值中间量 [%] / Kp deviation intermediate *)
    _fDti    : REAL;                         (* Ti 偏差中间量 [%] / Ti deviation intermediate *)
    _fDtd    : REAL;                         (* Td 偏差中间量 [%] / Td deviation intermediate *)
END_VAR
VAR CONSTANT
    DL_PDA_EPS    : REAL  := 1.0E-6;         (* 近零/容差判零容差（REAL 量级）[-] / Epsilon *)
    DL_PDA_CNTMAX : UDINT := 4294967295;     (* 计数饱和上限（R28）[-] / Count saturation cap *)
    DL_PDA_NMAX   : INT   := 100;            (* 确认拍数上限（防长时间不判）[拍] / Confirm scans cap *)
    c_fHun        : LREAL := 100.0;          (* 百分数换算常量（v1.0.1 由 VAR 迁入收口）[-] / Percent scale constant *)
END_VAR

(* —— 段 0：当拍判据派生 + 实例无条件刷新（R228A） —— *)
_bCfgBad := (fTolRel <= DL_PDA_EPS) OR (fTolAbs <= DL_PDA_EPS)                 (* 容差正域闸（两口径均须有效） / Tolerance gates *)
            OR (nConfirm < 1) OR (nConfirm > DL_PDA_NMAX);                     (* 确认拍数域闸 / Confirm-count gate *)
rtReset(CLK := bReset);                                                        (* 复位沿每拍必调 / Reset edge every scan *)
_bFinite := (fKp = fKp) AND ((fKp - fKp) = (fKp - fKp))                        (* Kp NaN 自反 + Inf 差判闸（v1.0.1）/ Kp NaN and Inf gates *)
            AND (fTi = fTi) AND ((fTi - fTi) = (fTi - fTi))                    (* Ti NaN 自反 + Inf 差判闸 / Ti NaN and Inf gates *)
            AND (fTd = fTd) AND ((fTd - fTd) = (fTd - fTd))                    (* Td NaN 自反 + Inf 差判闸 / Td NaN and Inf gates *)
            AND (fKpRef = fKpRef) AND ((fKpRef - fKpRef) = (fKpRef - fKpRef))  (* 基准 Kp NaN + Inf 闸 / Baseline Kp NaN and Inf gates *)
            AND (fTiRef = fTiRef) AND ((fTiRef - fTiRef) = (fTiRef - fTiRef))  (* 基准 Ti NaN + Inf 闸 / Baseline Ti NaN and Inf gates *)
            AND (fTdRef = fTdRef) AND ((fTdRef - fTdRef) = (fTdRef - fTdRef)); (* 基准 Td NaN + Inf 闸（Inf-Inf→NaN 漏报收口）/ Baseline Td NaN and Inf gates *)

(* —— 段 1：单拍量预清零（R107） —— *)
_bExKp := FALSE;                                                               (* Kp 越差预清 / Kp excursion preset *)
_bExTi := FALSE;                                                               (* Ti 越差预清 / Ti excursion preset *)
_bExTd := FALSE;                                                               (* Td 越差预清 / Td excursion preset *)
_bAny := FALSE;                                                                (* 汇总位预清 / Any preset *)
(* bDriftAny 不再每拍独立预清：改由段 5 由三确认位 OR 同源重算（v1.0.1，R52-06 汇总不回落） *)

(* —— 段 2：复位沿处理（作用域：清故障 + 清三个确认位 + 清计数 + 迁 eIdle，R283 逐项声明） —— *)
IF rtReset.Q THEN
    _bFault := FALSE;                                                          (* 清故障锁存 / Clear fault *)
    _eCause := E_DL_PdaCause.eNone;                                            (* 清成因 / Clear cause *)
    bDriftKp := FALSE;                                                         (* 清 Kp 确认位 / Clear Kp confirm *)
    bDriftTi := FALSE;                                                         (* 清 Ti 确认位 / Clear Ti confirm *)
    bDriftTd := FALSE;                                                         (* 清 Td 确认位 / Clear Td confirm *)
    nDriftCnt := 0;                                                            (* 清越差计数 / Clear count *)
    _nHold := 0;                                                               (* 清连续拍计数 / Clear hold counter *)
    fDriftKp := 0.0;                                                           (* 清 Kp 漂移出口 / Clear Kp drift outlet *)
    fDriftTi := 0.0;                                                           (* 清 Ti 漂移出口 / Clear Ti drift outlet *)
    fDriftTd := 0.0;                                                           (* 清 Td 漂移出口 / Clear Td drift outlet *)
    _eState := E_DL_PdaState.eIdle;                                            (* 迁未使能相 / Back to idle *)
END_IF

(* —— 段 3：组态故障锁存（锁存至复位沿，R189） —— *)
IF _bCfgBad AND NOT _bFault THEN
    _bFault := TRUE;                                                           (* 锁存故障位 / Latch fault *)
    _eCause := E_DL_PdaCause.eCfgIllegal;                                      (* 成因：组态非法 / Cause: illegal config *)
    _eState := E_DL_PdaState.eFault;                                           (* 同步迁故障相 / Migrate to fault *)
END_IF

(* —— 段 4：CASE 主状态机（ELSE 兜底迁 eFault，红线 6） —— *)
CASE _eState OF
    E_DL_PdaState.eIdle:                                                       (* 未使能：不审计，出口保持 / Disabled *)
        _nHold := 0;                                                           (* 失能清连续计数（防隐性回夹） / Clear hold *)
        IF bEnable AND NOT _bFault THEN
            _eState := E_DL_PdaState.eAudit;                                   (* 使能进入审计 / Enter audit *)
        END_IF
    E_DL_PdaState.eAudit:                                                      (* 审计相：三参数双口径比对 / Auditing *)
        IF NOT bEnable THEN
            _eState := E_DL_PdaState.eIdle;                                    (* 失能回未使能 / Back to idle *)
        ELSIF _bFinite THEN
            IF ABS(fKpRef) > DL_PDA_EPS THEN
                _fDkp := LREAL_TO_REAL(ABS(fKp - fKpRef) / ABS(fKpRef) * c_fHun);   (* 相对漂移 %：除子已过闸，显式窄化转换 / Relative drift, divisor gated *)
                _bExKp := _fDkp > LREAL_TO_REAL(fTolRel * c_fHun);             (* 越差判据：相对口径 / Excursion, relative *)
            ELSE
                _fDkp := ABS(fKp - fKpRef);                                    (* 基准近零：退化为绝对差（边界①） / Near-zero baseline: absolute *)
                _bExKp := _fDkp > fTolAbs;                                     (* 越差判据：绝对口径 / Excursion, absolute *)
            END_IF
            IF ABS(fTiRef) > DL_PDA_EPS THEN
                _fDti := LREAL_TO_REAL(ABS(fTi - fTiRef) / ABS(fTiRef) * c_fHun);   (* Ti 相对漂移 % / Ti relative drift *)
                _bExTi := _fDti > LREAL_TO_REAL(fTolRel * c_fHun);             (* Ti 越差判据 / Ti excursion *)
            ELSE
                _fDti := ABS(fTi - fTiRef);                                    (* Ti 基准为 0：绝对差（P 模式常见） / Ti near-zero: absolute *)
                _bExTi := _fDti > fTolAbs;                                     (* Ti 越差判据（绝对） / Ti excursion, absolute *)
            END_IF
            IF ABS(fTdRef) > DL_PDA_EPS THEN
                _fDtd := LREAL_TO_REAL(ABS(fTd - fTdRef) / ABS(fTdRef) * c_fHun);   (* Td 相对漂移 % / Td relative drift *)
                _bExTd := _fDtd > LREAL_TO_REAL(fTolRel * c_fHun);             (* Td 越差判据 / Td excursion *)
            ELSE
                _fDtd := ABS(fTd - fTdRef);                                    (* Td 基准为 0：绝对差 / Td near-zero: absolute *)
                _bExTd := _fDtd > fTolAbs;                                     (* Td 越差判据（绝对） / Td excursion, absolute *)
            END_IF
            fDriftKp := _fDkp;                                                 (* Kp 漂移出口（实时派生） / Kp drift outlet *)
            fDriftTi := _fDti;                                                 (* Ti 漂移出口 / Ti drift outlet *)
            fDriftTd := _fDtd;                                                 (* Td 漂移出口 / Td drift outlet *)
            _bAny := _bExKp OR _bExTi OR _bExTd;                               (* 任一越差汇总 / Any excursion *)
            IF _bAny THEN
                _nHold := _nHold + 1;                                          (* 连续越差拍递增 / Increment hold *)
            ELSE
                _nHold := 0;                                                   (* 有拍未越差即清零（降抖） / Reset on clean scan *)
            END_IF
            IF _nHold >= nConfirm THEN                                         (* 连续确认拍数到齐 / Confirm reached *)
                IF _bExKp THEN
                    bDriftKp := TRUE;                                          (* Kp 确认位锁存 / Latch Kp confirm *)
                END_IF
                IF _bExTi THEN
                    bDriftTi := TRUE;                                          (* Ti 确认位锁存 / Latch Ti confirm *)
                END_IF
                IF _bExTd THEN
                    bDriftTd := TRUE;                                          (* Td 确认位锁存 / Latch Td confirm *)
                END_IF
                IF nDriftCnt < DL_PDA_CNTMAX THEN
                    nDriftCnt := nDriftCnt + 1;                                (* 越差事件净额 +1（同拍多次不叠加） / Net +1 per confirmed event *)
                END_IF
                _nHold := 0;                                                   (* 计数归零，下一轮重新累积 / Restart accumulation *)
            END_IF
        END_IF                                                                 (* 非有限参数：本拍不判（保留确认位） / Non-finite: skip verdict *)
    E_DL_PdaState.eFault:                                                      (* 故障相：冻结保持末值，仅复位沿出 / Fault *)
        ;                                                                      (* 锁存回放（R28） / Replay from latch *)
    ELSE                                                                       (* 非法相位兜底迁安全态 / Illegal phase fallback *)
        _eState := E_DL_PdaState.eFault;                                       (* 迁故障相 / To fault *)
        _bFault := TRUE;                                                       (* 同步锁存 / Latch *)
        _eCause := E_DL_PdaCause.ePhaseBad;                                    (* 成因：非法相位 / Cause: illegal phase *)
END_CASE

(* —— 段 5：出口映射（bError/eState 同源，R191；bDriftAny 由三确认位 OR 同源重算，v1.0.1） —— *)
bDriftAny := bDriftKp OR bDriftTi OR bDriftTd;                                 (* 汇总出口同源重算（非有限拍不回落） / Any outlet re-derived *)
bError := _bFault;                                                             (* 故障标志镜像 / Fault flag mirror *)
eState := _eState;                                                             (* 状态出口 / State outlet *)
eCause := _eCause;                                                             (* 成因出口 / Cause outlet *)
END_FUNCTION_BLOCK

(* ---- FB_DL_PidParamGuard.st ---- *)
(*
  ==================================================================
  组件名 Component  : FB_DL_PidParamGuard
  分类   Category   : DL_Algo
  前缀   Naming     : FB_DL_ ｜ b/n/u/f/t/e/st 类型前缀制（R265）
  复杂度 Complexity  : 中
  版本   Version    : 1.0.0
  功能   Purpose    : PID 参数组在线运行期守卫（Kp/Ti/Td 有限性 + 域闸 + 退化降级）。
  来源   Source     : self-std（PID 参数治理公开语义自研）
  平台   Platform   : 纯 IEC 61131-3（比较 / ABS / R_TRIG），三平台通用
  分工声明 Split     : 与 FB_DL_PidParamDriftAudit 分工声明（R216）：本件做在线
                      参数闸（每拍有限性 + 域闸 + 退化降级，运行期保护）；后者
                      做离线漂移审计（趋势记录与慢漂分析）。两件双向互引，不
                      重复对方职责。
  作者   Author     : 道莅代码库 · PLC 编程专家（R61）
  归属 Ownership     : 本件无 TYPE 声明；引用件类型全部 IEC 标准原生。
  ------------------------------------------------------------------
  边界 Boundary     :
                      一 非有限入参 → 故障锁存 + 冻结上次合法快照（R187），
                         复位沿解除（bReset 恒可达，R152 自证）；
                      二 参数越界降级为上次合法值快照（不静默清零，R191 声明行：
                         bDegraded = TRUE + 出口保持快照），置信息级码；
                      三 快照更新只在「全部参数合法且域内」拍执行（保持槽写前
                         过闸，FB32-7）；首拍无快照时以域中点常量兜底（FB32-3
                         两级回退第二级）；
                      四 域闸上界须 > 下界（组态闸，逐对判，非法锁存同故障码）；
                      五 非有限闸逐个点名 9 个浮点入参（R272 全量枚举：fKp /
                         fTi / fTd / 六个域界引脚）；
                      六 无全局、无外部变量、无物理地址。
  错误码   Codes    :
    16#0002_3733【故障级】参数组含非有限值或域界组态非法，冻结快照，锁存至复位沿
    16#0002_3734【信息级】参数越域，已降级为上次合法快照（逐拍重算）
  验收   Acceptance :
    算法已证（脚本）：未跑 ｜ 编译器已证（三平台）：未跑
    V1 合法参数 → 三出口等于入参、bDegraded=FALSE
    V2 fKp=NaN → 码 3733、出口保持上次快照、锁存待复位
    V3 fKp 越上界 → 码 3734、fKpUse=上次快照、bDegraded=TRUE
  修订记录 Revision  :
    2026-11-21  v1.0.0  R61 首版（批 3 · 序号 11）
  ==================================================================
*)
FUNCTION_BLOCK FB_DL_PidParamGuard
VAR_INPUT
    bEnable : BOOL := TRUE;  // 使能，FALSE 时冻结快照出口（R191 声明行）/ the enable, false freezes the snapshot outlet
    bReset  : BOOL := FALSE; // 故障复位电平，上升沿清锁存 / the fault reset level
    fKp     : LREAL := 1.0;  // 比例增益入参 [-] / the proportional gain input
    fTi     : LREAL := 1.0;  // 积分时间入参 [秒] / the integral time input
    fTd     : LREAL := 0.0;  // 微分时间入参 [秒] / the derivative time input
    fKpMin  : LREAL := 0.0;  // 比例域下界 [-] / the proportional domain floor
    fKpMax  : LREAL := 100.0; // 比例域上界 [-] / the proportional domain ceiling
    fTiMin  : LREAL := 0.001; // 积分域下界 [秒] / the integral domain floor
    fTiMax  : LREAL := 3600.0; // 积分域上界 [秒] / the integral domain ceiling
    fTdMin  : LREAL := 0.0;  // 微分域下界 [秒] / the derivative domain floor
    fTdMax  : LREAL := 60.0; // 微分域上界 [秒] / the derivative domain ceiling
END_VAR
VAR_OUTPUT
    fKpUse    : LREAL := 1.0;  // 比例增益出口（快照或原值）[-] / the proportional gain outlet
    fTiUse    : LREAL := 1.0;  // 积分时间出口 [秒] / the integral time outlet
    fTdUse    : LREAL := 0.0;  // 微分时间出口 [秒] / the derivative time outlet
    bDegraded : BOOL := FALSE; // 本拍降级标志（信息级伴随）[-] / the degraded flag of this scan
    bError    : BOOL := FALSE; // 故障锁存位（与锁存同源，R191）/ the fault bit from the latch
    bValid    : BOOL := FALSE; // 参数可用标志 [-] / the parameters usable flag
    eErr      : UDINT := 16#0000_0000; // 错误码，0 = 正常 / the error code, zero is ok
END_VAR
VAR
    _bInit    : BOOL := FALSE; // 首拍初始化标志（R310）/ the first scan flag
    _bFault   : BOOL := FALSE; // 故障锁存副本（仅复位沿清除）/ the fault latch copy
    _bFin     : BOOL := FALSE; // 非有限闸结果（逐拍重算）/ the finiteness gate result
    _bInDom   : BOOL := FALSE; // 域闸结果（逐拍重算）/ the domain gate result
    _bDomCfg  : BOOL := FALSE; // 域界组态合法标记（逐拍重算）/ the domain configuration flag
    _fKpSnap  : LREAL := 1.0;  // 比例快照（仅合法拍更新）/ the proportional snapshot
    _fTiSnap  : LREAL := 1.0;  // 积分快照 / the integral snapshot
    _fTdSnap  : LREAL := 0.0;  // 微分快照 / the derivative snapshot
    rtReset   : R_TRIG; // 复位沿实例，段 0 无条件刷新 / the reset edge instance
END_VAR

// 段 0｜复位沿无条件周期刷新（禁入分支，R7）/ segment 0, the unconditional refresh
rtReset(CLK := bReset); // 复位沿 / the reset edge

// 段 1｜首拍初始化与复位沿作用域（R310 / R311）/ segment 1, the first scan init and the reset scope
IF NOT _bInit THEN // 首拍一拍 / the first scan
    _bInit := TRUE; // 置首拍标志 / raise the first scan flag
    _bFault := FALSE; // 故障锁存显式清零 / clear the fault latch explicitly
    _fKpSnap := fKp; // 首拍以入参装快照（入参缺省即域内默认）/ seed the snapshot from the input
    _fTiSnap := fTi; // 积分快照装填 / seed the integral snapshot
    _fTdSnap := fTd; // 微分快照装填 / seed the derivative snapshot
END_IF
IF rtReset.Q THEN // 复位沿（作用域：仅清锁存，快照保持最近合法值，R311 声明）/ the reset edge clears the latch only
    _bFault := FALSE; // 清故障锁存（解除路径：复位沿恒可达，R152 自证）/ clear the fault latch
END_IF

// 段 2｜非有限闸：9 个浮点入参逐个点名（R272 全量，边界五）/ segment 2, the finiteness gate naming all nine floating pins
_bFin := (fKp = fKp) AND ((fKp - fKp) = (fKp - fKp))
AND (fTi = fTi) AND ((fTi - fTi) = (fTi - fTi))
AND (fTd = fTd) AND ((fTd - fTd) = (fTd - fTd))
AND (fKpMin = fKpMin) AND ((fKpMin - fKpMin) = (fKpMin - fKpMin))
AND (fKpMax = fKpMax) AND ((fKpMax - fKpMax) = (fKpMax - fKpMax))
AND (fTiMin = fTiMin) AND ((fTiMin - fTiMin) = (fTiMin - fTiMin))
AND (fTiMax = fTiMax) AND ((fTiMax - fTiMax) = (fTiMax - fTiMax))
AND (fTdMin = fTdMin) AND ((fTdMin - fTdMin) = (fTdMin - fTdMin))
AND (fTdMax = fTdMax) AND ((fTdMax - fTdMax) = (fTdMax - fTdMax)); // NaN 自反 + Inf 差值自减逐项 / the reflexive and difference tests term by term

// 段 3｜域界组态闸与域闸（边界四）/ segment 3, the domain configuration and the domain gates
_bDomCfg := (fKpMax > fKpMin) AND (fTiMax > fTiMin) AND (fTdMax > fTdMin); // 三对域界严格递增 / the three strictly increasing pairs
_bInDom := (fKp >= fKpMin) AND (fKp <= fKpMax)
AND (fTi >= fTiMin) AND (fTi <= fTiMax)
AND (fTd >= fTdMin) AND (fTd <= fTdMax); // 三参数域内判 / the three parameters inside the domains
IF (NOT _bFin) OR (NOT _bDomCfg) THEN // 非有限或域界非法：故障锁存（边界一）/ a non finite or an illegal domain configuration
    _bFault := TRUE; // 锁存故障（3733，出口回放）/ latch the fault
END_IF

// 段 4｜快照闸与降级（边界二三）/ segment 4, the snapshot gate and the degradation
IF _bFin AND _bDomCfg AND _bInDom THEN // 全部合法：出口 = 原值并更新快照（保持槽写前过闸，FB32-7）/ all legal, the outlet takes the values and updates the snapshot
    _fKpSnap := fKp; // 快照更新 / update the snapshot
    _fTiSnap := fTi; // 快照更新 / update the snapshot
    _fTdSnap := fTd; // 快照更新 / update the snapshot
    bDegraded := FALSE; // 无降级 / no degradation
ELSIF (NOT _bFault) THEN // 域外但无锁存：降级为快照（不静默清零，边界二）/ out of the domain without a latch, degrade to the snapshot
    bDegraded := TRUE; // 置降级标志 / raise the degraded flag
ELSE // 故障锁存态：出口冻结快照（R191 声明行）/ the latched state freezes the snapshot outlet
    bDegraded := FALSE; // 降级标志不置（故障码已表达）/ the degraded flag stays low
END_IF

// 段 5｜统一出口（冻结语义：保持上次合法快照，R191 / R273 防污染：快照本身写前过闸）/ segment 5, the unified outlet
fKpUse := _fKpSnap; // 比例出口 / the proportional outlet
fTiUse := _fTiSnap; // 积分出口 / the integral outlet
fTdUse := _fTdSnap; // 微分出口 / the derivative outlet
bError := _bFault; // 故障位出口（与锁存同源）/ the fault bit outlet
bValid := (NOT _bFault) AND (NOT bDegraded); // 参数可用标志 / the usable flag
IF _bFault THEN // 故障锁存回放（R187）/ the latched fault replays
    eErr := 16#0002_3733; // 故障级：参数非有限或域界组态非法 / fault grade, the non finite parameter or the illegal domain
ELSIF bDegraded THEN // 降级（信息级不置 bError，R285 口径）/ the degraded informational code
    eErr := 16#0002_3734; // 信息级：参数越域已降级为快照 / informational, degraded to the snapshot
ELSE // 无事件 / no event
    eErr := 16#0000_0000; // 正常 / ok
END_IF
END_FUNCTION_BLOCK

(* ---- FB_DL_PidRelayAutoTune.st ---- *)
(*
  Name        : FB_DL_PidRelayAutoTune
  Category    : DL_Algo
  Version     : 1.0.0
  Purpose     : 继电器反馈自整定：强制振荡观测极限周期/幅值，按 Åström-Hägglund 公开公式给 PID 初值（Kp = 4d/πa，Ti = Tu/2，Td = Tu/8）；/ Relay-feedback auto-tuning: forced-oscillation observation of ultimate period and amplitude, PID seed values from the published Astrom-Hagglund formulas
  溯源        : 自研-公开方法（relay-tuning 公开公式），clean-room 实现
  Boundary    : ① 迟滞带宽/激励幅值/采样周期三重正域闸，任一越域锁存故障；
                ② 振荡周期须测得 ≥ 3 个完整周期且逐周期稳定才出参数（防半波截断算错极限周期）；
                ③ 出口 PID 初值域钳位（Kp > 0、Ti > 0、Td >= 0），幅值发散或周期不稳 → 有效性出口 FALSE 且不出参数；
                ④ 整定中不写控制输出：本件零控制量引脚，仅出继电器建议态信号（属主边界，防误动作）；
                ⑤ 非有限测量该拍不入振荡检测（计时暂停非快进，防污染周期窗）；
                ⑥ 超时未达成 3 周期为信息级（不置故障标志，成因出口可查）。
*)
TYPE E_DL_PatState :
(
    eIdle  := 0,                             (* 未整定 / Not tuning *)
    eRelay := 10,                            (* 继电器振荡观测中 / Relay oscillation observing *)
    eReady := 20,                            (* 整定完成（有效性查 bValid 出口） / Tuning finished, see bValid *)
    eFault := 90                             (* 故障锁存相 / Fault latched *)
);
END_TYPE

TYPE E_DL_PatCause :
(
    eNone      := 0,                         (* 无成因 / No cause *)
    eCfgIllegal:= 1,                        (* 组态非法：幅值/迟滞/周期越域 / Illegal config *)
    eNoOsc     := 2,                        (* 信息级：未达成 3 稳定周期（超时/发散） / Info: no stable periods *)
    ePhaseBad  := 3                         (* 非法相位兜底 / Illegal phase fallback *)
);
END_TYPE

FUNCTION_BLOCK FB_DL_PidRelayAutoTune
VAR_INPUT
    fMeas    : REAL := 0.0;                  (* 被整定回路测量值（任意工程量）[-] / Loop measurement *)
    fSetpoint: REAL := 50.0;                 (* 振荡基准（被控量目标中值）[-] / Oscillation reference *)
    fRelayAmp: REAL := 5.0;                  (* 继电器激励幅值，域 > 0 [工程单位] / Relay excitation amplitude *)
    fHyst    : REAL := 1.0;                  (* 迟滞半带宽，域 > 0 且 < 幅值 [工程单位] / Hysteresis half band *)
    tSample  : TIME := T#100MS;              (* 采样周期，域 > T#0S [ms] / Sampling period *)
    tWatch   : TIME := T#120S;               (* 整定观测总超时，域 > T#0S [ms] / Tuning watch timeout *)
    bStart   : BOOL := FALSE;                (* 启动整定命令，上升沿进入观测 [-] / Start tuning command *)
    bEnable  : BOOL := TRUE;                 (* 使能 [-] / Enable *)
    bReset   : BOOL := FALSE;                (* 复位命令，上升沿清故障与结果 [-] / Reset command *)
END_VAR
VAR_OUTPUT
    bRelaySug: BOOL;                         (* 继电器建议态（属主自行施加，本件不写控制输出）[-] / Suggested relay state *)
    nCycles  : INT;                          (* 已测得完整周期数 [个] / Complete periods measured *)
    fKp      : REAL;                         (* PID 初值：比例增益 [-] / PID seed: gain *)
    fTi      : REAL;                         (* PID 初值：积分时间 [s] / PID seed: integral time *)
    fTd      : REAL;                         (* PID 初值：微分时间 [s] / PID seed: derivative time *)
    bValid   : BOOL;                         (* 参数有效性出口（3 稳定周期达成才 TRUE）[-] / Parameter validity *)
    eState   : E_DL_PatState;                (* 状态出口 / State outlet *)
    eCause   : E_DL_PatCause;                (* 成因出口（R190 归因唯一） / Cause outlet *)
    bError   : BOOL;                         (* 故障锁存标志 [-] / Fault latch flag *)
END_VAR
VAR
    _eState : E_DL_PatState := E_DL_PatState.eIdle;  (* 内部相位（CASE 唯一写入目标） / Internal phase *)
    _eCause : E_DL_PatCause := E_DL_PatCause.eNone;  (* 成因锁存量 / Latched cause *)
    rtStart : R_TRIG;                        (* 启动沿实例，段 0 无条件调用 / Start edge instance *)
    rtReset : R_TRIG;                        (* 复位沿实例，段 0 无条件调用 / Reset edge instance *)
    _bFault : BOOL;                          (* 故障锁存位 / Latched fault bit *)
    _bCfgBad: BOOL;                          (* 组态非法当拍量 / Illegal config this scan *)
    _bFin   : BOOL;                          (* 测量有限性当拍量 / Measurement finiteness *)
    _bRelayI: BOOL;                          (* 继电器态内部量（迟滞保持）[-] / Relay state internal *)
    _bPrevRel: BOOL;                         (* 上拍继电器态（沿检测）[-] / Previous relay state *)
    _bUpCr  : BOOL;                          (* 本拍向上穿越当拍量（继电器态由高变低）[-] / Upward crossing this scan *)
    _fDtSec : REAL;                          (* 采样周期秒值，域 > eps [s] / Sampling period seconds *)
    _fTacc  : REAL;                          (* 周期计时累加量 [s] / Period time accumulator *)
    _fTune  : REAL;                          (* 整定总耗时累加量 [s] / Total tuning elapsed *)
    _fTu1   : REAL;                          (* 周期样本 1 [s] / Period sample 1 *)
    _fTu2   : REAL;                          (* 周期样本 2 [s] / Period sample 2 *)
    _fTu3   : REAL;                          (* 周期样本 3 [s] / Period sample 3 *)
    _nTuN   : INT;                           (* 已存周期样本数 [个] / Stored period samples *)
    _fPk    : REAL;                          (* 本周期峰值 [工程单位] / Cycle peak *)
    _fTr    : REAL;                          (* 本周期谷值 [工程单位] / Cycle trough *)
    _fAmp   : REAL;                          (* 上周期振荡半幅值 [工程单位] / Previous cycle amplitude *)
    _fAmI   : REAL;                          (* 本周期半幅值中间量 [工程单位] / Current amplitude *)
    _fKpI   : REAL;                          (* Kp 中间量（出参域钳前）[-] / Kp intermediate *)
    _fTiI   : REAL;                          (* Ti 中间量 [s] / Ti intermediate *)
    _fTdI   : REAL;                          (* Td 中间量 [s] / Td intermediate *)
END_VAR
VAR CONSTANT
    DL_PAT_EPS   : REAL := 1.0E-6;           (* 判零容差 [-] / Epsilon *)
    DL_PAT_PI    : REAL := 3.14159265;       (* 圆周率常量（公开公式用）[-] / Pi constant *)
    DL_PAT_TUSTAB: REAL := 0.2;              (* 周期稳定相对容差（20%）[-] / Period stability tolerance *)
    DL_PAT_AMPDIV: REAL := 0.5;              (* 幅值发散相对判据（50%）[-] / Amplitude divergence ratio *)
    DL_PAT_NNEED : INT   := 3;               (* 完整周期需求数（边界②）[个] / Required periods *)
END_VAR

(* —— 段 0：当拍判据派生 + 实例无条件刷新（R228A） —— *)
_fDtSec := TIME_TO_LREAL(tSample) / 1000.0;              (* 采样周期秒化（除子常量 1000） / Period seconds *)
_bCfgBad := (fRelayAmp <= DL_PAT_EPS) OR (fHyst <= DL_PAT_EPS) OR (fHyst >= fRelayAmp)   (* 幅值/迟滞正域闸（边界①） / Amplitude and hysteresis gates *)
            OR NOT (tSample > T#0S) OR NOT (tWatch > T#0S);   (* 采样/超时周期正域闸（边界①） / Period gates *)
rtStart(CLK := bStart);                                  (* 启动沿每拍必调 / Start edge every scan *)
rtReset(CLK := bReset);                                  (* 复位沿每拍必调 / Reset edge every scan *)
_bFin := (fMeas = fMeas) AND ((fMeas - fMeas) = (fMeas - fMeas));   (* 测量 NaN 自反 + Inf 差判闸 / Measurement NaN and Inf gate *)
_bUpCr := FALSE;                                         (* 向上穿越当拍量预清 / Crossing preset *)
_bPrevRel := _bRelayI;                                   (* 上拍继电器态快照 / Relay state snapshot *)

(* —— 段 1：单拍量预清零（R107） —— *)
bRelaySug := _bRelayI;                                   (* 建议态出口 = 内部保持量（确定值） / Suggested relay outlet *)

(* —— 段 2：复位沿处理（作用域：清故障 + 清结果 + 迁 eIdle，R283 逐项声明） —— *)
IF rtReset.Q THEN
    _bFault := FALSE;                                    (* 清故障锁存 / Clear fault *)
    _eCause := E_DL_PatCause.eNone;                      (* 清成因 / Clear cause *)
    bValid := FALSE;                                     (* 清有效性出口 / Clear validity *)
    fKp := 0.0; fTi := 0.0; fTd := 0.0;                  (* 清 PID 初值出口 / Clear PID seed outlets *)
    nCycles := 0;                                        (* 清周期数出口 / Clear cycles *)
    _nTuN := 0; _fTacc := 0.0; _fTune := 0.0;            (* 清样本数/计时/耗时 / Clear samples and timers *)
    _bRelayI := FALSE;                                   (* 清继电器态 / Clear relay state *)
    _eState := E_DL_PatState.eIdle;                      (* 迁未整定相 / Back to idle *)
END_IF

(* —— 段 3：组态故障锁存（锁存至复位沿，R189） —— *)
IF _bCfgBad AND NOT _bFault THEN
    _bFault := TRUE;                                     (* 锁存故障位 / Latch fault *)
    _eCause := E_DL_PatCause.eCfgIllegal;                (* 成因：组态非法 / Cause illegal config *)
    _eState := E_DL_PatState.eFault;                     (* 同步迁故障相 / Migrate to fault *)
END_IF

(* —— 段 4：CASE 主状态机（ELSE 兜底迁 eFault，红线 6） —— *)
CASE _eState OF
    E_DL_PatState.eIdle:                                 (* 未整定：出口保持确定值 / Idle *)
        bValid := FALSE;                                 (* 未整定有效性 FALSE（不留陈旧） / Validity false *)
        IF rtStart.Q AND bEnable AND NOT _bFault THEN
            _nTuN := 0; _fTacc := 0.0; _fTune := 0.0;    (* 清样本数/计时/耗时（新整定轮） / Clear samples and timers *)
            _fPk := fMeas; _fTr := fMeas;                (* 峰谷以首拍测量锚定 / Anchor peak and trough *)
            _fAmp := 0.0;                                (* 清上周期幅值 / Clear previous amplitude *)
            _bRelayI := FALSE;                           (* 继电器态从低起始 / Relay from low *)
            _eState := E_DL_PatState.eRelay;             (* 进入观测相 / Enter observing *)
        END_IF
    E_DL_PatState.eRelay:                                (* 观测相：迟滞继电器 + 周期/幅值测量 / Observing *)
        IF NOT bEnable THEN
            _eState := E_DL_PatState.eIdle;              (* 失能回未整定 / Back to idle *)
        ELSIF _bFin AND (_fDtSec > DL_PAT_EPS) THEN      (* 非有限拍整拍跳过（边界⑤） / Skip non-finite scan *)
            _fTacc := _fTacc + _fDtSec;                  (* 周期计时累加（暂停非快进） / Period acc advance *)
            _fTune := _fTune + _fDtSec;                  (* 总耗时累加 / Elapsed advance *)
            IF (NOT _bRelayI AND (fMeas < fSetpoint - fHyst)) OR (_bRelayI AND (fMeas > fSetpoint + fHyst)) THEN
                _bRelayI := NOT _bRelayI;                (* 迟滞带直比翻转（禁浮点等值） / Hysteresis band toggle *)
            END_IF
            IF _bPrevRel AND NOT _bRelayI THEN
                _bUpCr := TRUE;                          (* 向上穿越沿（低 → 高穿越上带） / Upward crossing edge *)
            END_IF
            IF fMeas > _fPk THEN
                _fPk := fMeas;                           (* 本周期峰值刷新 / Cycle peak update *)
            END_IF
            IF fMeas < _fTr THEN
                _fTr := fMeas;                           (* 本周期谷值刷新 / Cycle trough update *)
            END_IF
            IF _bUpCr THEN                               (* 向上穿越：收口一个完整周期 / Crossing closes a period *)
                IF _nTuN >= 1 THEN
                    IF _nTuN = 1 THEN
                        _fTu1 := _fTacc;                 (* 周期样本 1 收存 / Store sample 1 *)
                    ELSIF _nTuN = 2 THEN
                        _fTu2 := _fTacc;                 (* 周期样本 2 收存 / Store sample 2 *)
                    END_IF
                    _fAmp := _fAmI; _fAmI := (_fPk - _fTr) / 2.0;   (* 幅值转存 + 本周期半幅值（除子常量 2） / Amplitude roll *)
                END_IF
                _nTuN := _nTuN + 1;                      (* 完整周期计数净额 +1 / Period count *)
                IF _nTuN > 3 THEN _fTu3 := _fTacc; END_IF   (* 周期样本 3 收存（覆盖） / Store sample 3 *)
                _fTacc := 0.0;                           (* 周期计时重置（R227） / Period acc reset *)
                _fPk := fMeas; _fTr := fMeas;            (* 峰谷重锚定 / Peak and trough re-anchor *)
            END_IF
            IF (_fTu1 > DL_PAT_EPS) AND (_fTu2 > DL_PAT_EPS) AND (_fTu3 > DL_PAT_EPS) AND (_nTuN >= DL_PAT_NNEED + 1) THEN
                IF (ABS(_fTu3 - _fTu2) <= DL_PAT_TUSTAB * _fTu3) AND (ABS(_fTu2 - _fTu1) <= DL_PAT_TUSTAB * _fTu2) THEN
                    _fKpI := 4.0 * fRelayAmp / (DL_PAT_PI * _fAmI);   (* 周期稳定 + 公开公式 Kp（除子已过幅值正域闸，边界②③） / Stable periods, formula Kp *)
                    _fTiI := _fTu3 / 2.0;                (* 公开公式 Ti（除子常量 2） / Formula Ti *)
                    _fTdI := _fTu3 / 8.0;                (* 公开公式 Td（除子常量 8） / Formula Td *)
                    IF (_fAmI > DL_PAT_EPS) AND (_fKpI > 0.0) AND (_fTiI > 0.0) AND (_fTdI >= 0.0) THEN
                        fKp := _fKpI; fTi := _fTiI; fTd := _fTdI;   (* PID 初值出口（域钳后放行，边界③） / PID seed outlets *)
                        bValid := TRUE;                  (* 有效性 TRUE / Validity true *)
                        nCycles := _nTuN - 1;            (* 已测完整周期数出口 / Cycles outlet *)
                        _eState := E_DL_PatState.eReady; (* 迁整定完成相 / To ready *)
                    ELSE
                        bValid := FALSE; nCycles := _nTuN - 1;   (* 域钳拦截不出参数（边界③） / Clamp reject *)
                        _eCause := E_DL_PatCause.eNoOsc; (* 信息级成因（不置 bError，边界⑥） / Info cause *)
                        _eState := E_DL_PatState.eReady; (* 迁完成相（无效结论） / To ready invalid *)
                    END_IF
                ELSE
                    bValid := FALSE; nCycles := _nTuN - 1;   (* 周期不稳不出参数（边界③） / Unstable: invalid *)
                    _eCause := E_DL_PatCause.eNoOsc;     (* 信息级成因（边界⑥） / Info cause *)
                    _eState := E_DL_PatState.eReady;     (* 迁完成相（无效结论） / To ready invalid *)
                END_IF
            ELSIF _fTune > TIME_TO_LREAL(tWatch) THEN    (* 总超时：未达成 3 周期（信息级） / Watch timeout *)
                bValid := FALSE;                         (* 不出参数（边界②） / No parameters *)
                nCycles := _nTuN - 1;                    (* 已达成周期数照报 / Cycles outlet *)
                IF nCycles < 0 THEN nCycles := 0; END_IF (* 负数钳零（半周期不计） / Clamp negative *)
                _eCause := E_DL_PatCause.eNoOsc;         (* 信息级成因（边界⑥） / Info cause *)
                _eState := E_DL_PatState.eReady;         (* 迁完成相（无效结论） / To ready invalid *)
            END_IF
        END_IF
    E_DL_PatState.eReady:                                (* 完成相：结论与参数冻结保持 / Ready *)
        IF rtStart.Q THEN
            _eState := E_DL_PatState.eIdle;              (* 新启动沿经 eIdle 重入（防隐性回夹） / Restart via idle *)
        END_IF
    E_DL_PatState.eFault:                                (* 故障相：冻结保持，仅复位沿出 / Fault *)
        ;                                                (* 锁存回放（R28） / Replay from latch *)
    ELSE                                                 (* 非法相位兜底迁安全态 / Illegal phase fallback *)
        _eState := E_DL_PatState.eFault; _bFault := TRUE;   (* 迁故障相 + 同步锁存 / To fault and latch *)
        _eCause := E_DL_PatCause.ePhaseBad;              (* 成因：非法相位 / Cause illegal phase *)
END_CASE

(* —— 段 5：出口映射（bError/eState 同源，R191） —— *)
bRelaySug := _bRelayI;                                   (* 继电器建议态出口（观测相实时镜像） / Relay suggestion outlet *)
bError := _bFault;                                       (* 故障标志镜像 / Fault flag mirror *)
eState := _eState;                                       (* 状态出口 / State outlet *)
eCause := _eCause;                                       (* 成因出口 / Cause outlet *)
END_FUNCTION_BLOCK

(* ---- FB_DL_PumpSurgeGuard.st ---- *)
(*
  Name        : FB_DL_PumpSurgeGuard
  Category    : DL_Algo
  Version     : 1.0.0
  Purpose     : 泵喘振区逼近保护：以流量-压力工况点对线性喘振线求裕度，裕度低于门槛自动降载（流量上限限幅输出），恢复期斜坡回升；/ Pump surge guard: margin of the operating point against a linear surge line; below threshold the flow setpoint is automatically derated and ramped back on recovery
  溯源        : 借 t1-1-oscat-basic ◐/自研 的分类/参数域组织，clean-room 实现
  Boundary    : ① 组态闸：流量量程/裕度门槛/斜坡速率/周期任一越域或裕度门槛 > 1 → 锁存故障（量程 0 使裕度无定义）；
                ② 除零前置：流量上限比除子为 fFlowCmd，仅 |fFlowCmd| > eps 时计算（流量命令近零视为已充分降载，斜坡目标取 1）；
                ③ 非有限流量/压力该拍不更新判据（斜坡保持上拍值，防污染降载器）；
                ④ 裕度与降载系数均饱和 0..1，饱和是该变量最后一次写；
                ⑤ 降载斜坡按 fRampRate（1/s）× 周期秒值逐拍逼近目标，无突跳；
                ⑥ 本件为保护层，只限幅不切泵（启停由上层顺序控制，属主边界）。
*)
TYPE E_DL_PsgState :
(
    eIdle  := 0,                             (* 未使能 / Disabled *)
    eRun   := 10,                            (* 喘振保护运行 / Guarding *)
    eFault := 90                             (* 故障锁存相 / Fault latched *)
);
END_TYPE

TYPE E_DL_PsgCause :
(
    eNone       := 0,                        (* 无故障成因 / No cause *)
    eCfgIllegal := 1,                        (* 组态非法：量程/门槛/斜坡越域 / Illegal config *)
    eSurge      := 2,                        (* 裕度低于门槛（降载激活） / Margin below threshold *)
    ePhaseBad   := 3                         (* 非法相位兜底 / Illegal phase fallback *)
);
END_TYPE

FUNCTION_BLOCK FB_DL_PumpSurgeGuard
VAR_INPUT
    fFlow      : REAL := 0.0;                (* 泵流量实测 [m3/h] / Measured pump flow *)
    fPress     : REAL := 0.0;                (* 泵出口压力实测（扬程口径）[bar] / Measured discharge pressure *)
    fFlowCmd   : REAL := 0.0;                (* 上层流量设定（降载比基准）[m3/h] / Upstream flow setpoint *)
    fPressRef  : REAL := 5.0;               (* 喘振线参考压力（线截距基准），域 >= 0 [bar] / Surge-line reference pressure *)
    fSlope     : REAL := 0.2;                (* 喘振线斜率（压升 1 bar 对应喘振流量下限增量），域 >= 0 [(m3/h)/bar] / Surge-line slope *)
    fFlowSpan  : REAL := 100.0;              (* 流量量程（裕度归一化分母），域 > 0 [m3/h] / Flow span for margin normalisation *)
    fMarginMin : REAL := 0.15;               (* 裕度门槛（低于即降载），域 (0..1] [-] / Margin threshold, (0..1] *)
    fRampRate  : REAL := 0.1;               (* 降载/恢复斜坡速率，域 > 0 [1/s] / Ramp rate, > 0 *)
    tCycle     : TIME := T#100MS;           (* 运行周期，域 > T#0S [ms] / Cycle period, > 0 *)
    bEnable    : BOOL := TRUE;              (* 保护使能 [-] / Enable *)
    bReset     : BOOL := FALSE;             (* 复位命令，上升沿清降载与故障 [-] / Reset command *)
END_VAR
VAR_OUTPUT
    fMargin    : REAL;                      (* 工况点距喘振线归一化裕度 0..1（饱和）[-] / Normalised surge margin, saturated *)
    fFlowLimit : REAL;                      (* 降载后流量上限（fFlowCmd × 系数）[m3/h] / Derated flow limit *)
    fDerateFac : REAL;                      (* 降载系数 0..1（斜坡逼近）[-] / Derating factor, ramped *)
    bSurgeWarn : BOOL;                      (* 喘振逼近告警（裕度 < 门槛，电平）[-] / Surge proximity warning *)
    eState     : E_DL_PsgState;             (* 状态出口 / State outlet *)
    eCause     : E_DL_PsgCause;             (* 故障成因出口（R190 归因唯一） / Fault cause outlet *)
    bError     : BOOL;                      (* 故障锁存标志 [-] / Fault latch flag *)
END_VAR
VAR
    _eState   : E_DL_PsgState := E_DL_PsgState.eIdle;    (* 内部相位（CASE 唯一写入目标） / Internal phase *)
    _eCause   : E_DL_PsgCause := E_DL_PsgCause.eNone;    (* 故障成因锁存量 / Latched cause *)
    rtReset   : R_TRIG;                       (* 复位沿实例，段 0 无条件调用 / Reset edge instance *)
    _bFault   : BOOL;                         (* 故障锁存位 / Latched fault bit *)
    _bCfgBad  : BOOL;                         (* 组态非法当拍量 / Illegal config this scan *)
    _bFin     : BOOL;                         (* 输入有限性当拍量（流量/压力联合） / Input finiteness joint *)
    _fDtSec   : REAL;                         (* 周期折算秒值，域 > eps [s] / Period in seconds *)
    _fSurgeFl : REAL;                         (* 当前压力下喘振流量下限 [m3/h] / Surge flow limit at pressure *)
    _fMargI   : REAL;                         (* 裕度中间量（饱和前）[-] / Margin intermediate *)
    _fTarget  : REAL;                         (* 降载系数斜坡目标 [-] / Derating ramp target *)
    _fStep    : REAL;                         (* 本拍斜坡步长 [1/s 口径] / Ramp step this scan *)
    _fFac     : REAL;                         (* 降载系数内部量 0..1 [-] / Derating factor internal *)
END_VAR
VAR CONSTANT
    DL_PSG_EPS    : REAL := 1.0E-6;           (* 判零容差 [-] / Epsilon *)
    DL_PSG_PCTMAX : REAL := 1.0;              (* 裕度/系数满量程（归一化上限）[-] / Full scale *)
    DL_PSG_PCTMIN : REAL := 0.0;              (* 裕度/系数下限 [-] / Lower bound *)
    DL_PSG_DERMAX : REAL := 0.4;              (* 降载系数下限（最多降到 40%，防深喘振区反复进出）[-] / Derating floor *)
END_VAR

(* —— 段 0：当拍判据派生 + 实例无条件刷新（R228A） —— *)
_fDtSec := TIME_TO_LREAL(tCycle) / 1000.0;                                     (* 周期秒化（除子常量 1000） / Period to seconds *)
_bCfgBad := NOT (tCycle > T#0S)                                                (* 周期正域闸 / Period gate *)
            OR (fFlowSpan <= DL_PSG_EPS)                                       (* 流量量程正域闸（裕度除子） / Flow span gate *)
            OR (fPressRef < 0.0) OR (fSlope < 0.0)                             (* 参考压力/斜率非负闸 / Reference and slope gates *)
            OR (fMarginMin <= DL_PSG_EPS) OR (fMarginMin > DL_PSG_PCTMAX)      (* 裕度门槛域闸 (0..1] / Margin threshold gate *)
            OR (fRampRate <= DL_PSG_EPS);                                      (* 斜坡速率正域闸 / Ramp rate gate *)
rtReset(CLK := bReset);                                                        (* 复位沿每拍必调 / Reset edge every scan *)
_bFin := (fFlow = fFlow) AND (fPress = fPress)                                 (* 流量/压力 NaN 自反闸 / Flow and pressure NaN gates *)
            AND ((fFlow - fFlow) = (fFlow - fFlow))                            (* 流量 Inf 差判闸 / Flow Inf gate *)
            AND ((fPress - fPress) = (fPress - fPress));                       (* 压力 Inf 差判闸 / Pressure Inf gate *)

(* —— 段 1：单拍量预清零（R107；fDerateFac 为斜坡状态量，不在此预清） —— *)
fMargin := 0.0;                                                                (* 裕度出口预清 / Margin outlet preset *)
bSurgeWarn := FALSE;                                                           (* 告警出口预清 / Warn outlet preset *)
_fMargI := 0.0;                                                                (* 裕度中间量预置（非有限拍保持 0 语义） / Margin intermediate preset *)
_fTarget := DL_PSG_PCTMAX;                                                     (* 斜坡目标预置（默认全流量） / Ramp target preset *)

(* —— 段 2：复位沿处理（作用域：清故障 + 清降载系数与限幅 + 迁 eIdle，R283 逐项声明） —— *)
IF rtReset.Q THEN
    _bFault := FALSE;                                                          (* 清故障锁存 / Clear fault *)
    _eCause := E_DL_PsgCause.eNone;                                            (* 清成因 / Clear cause *)
    _fFac := DL_PSG_PCTMAX;                                                    (* 降载系数回 1（不降载） / Factor back to 1 *)
    fDerateFac := DL_PSG_PCTMAX;                                               (* 系数出口回 1 / Factor outlet back to 1 *)
    fFlowLimit := 0.0;                                                         (* 清限幅出口 / Clear limit outlet *)
    _eState := E_DL_PsgState.eIdle;                                            (* 迁未使能相 / Back to idle *)
END_IF

(* —— 段 3：组态故障锁存（锁存至复位沿，R189） —— *)
IF _bCfgBad AND NOT _bFault THEN
    _bFault := TRUE;                                                           (* 锁存故障位 / Latch fault *)
    _eCause := E_DL_PsgCause.eCfgIllegal;                                      (* 成因：组态非法 / Cause: illegal config *)
    _eState := E_DL_PsgState.eFault;                                           (* 同步迁故障相 / Migrate to fault *)
END_IF

(* —— 段 4：CASE 主状态机（ELSE 兜底迁 eFault，红线 6） —— *)
CASE _eState OF
    E_DL_PsgState.eIdle:                                                       (* 未使能：不保护，出口确定值 / Disabled *)
        fMargin := 0.0;                                                        (* 失能清裕度出口 / Clear margin outlet *)
        bSurgeWarn := FALSE;                                                   (* 失能清告警出口 / Clear warn outlet *)
        fFlowLimit := 0.0;                                                     (* 失能清限幅出口 / Clear limit outlet *)
        fDerateFac := DL_PSG_PCTMAX;                                           (* 失能系数回 1（不降载语义） / Factor outlet back to 1 *)
        _fFac := DL_PSG_PCTMAX;                                                (* 内部系数同步回 1 / Internal factor reset *)
        IF bEnable AND NOT _bFault THEN
            _eState := E_DL_PsgState.eRun;                                     (* 使能进入保护 / Enter guarding *)
        END_IF
    E_DL_PsgState.eRun:                                                        (* 保护相：裕度判据 + 斜坡降载 / Guarding *)
        IF NOT bEnable THEN
            _eState := E_DL_PsgState.eIdle;                                    (* 失能回未使能 / Back to idle *)
        ELSIF _bFin AND (_fDtSec > DL_PSG_EPS) THEN
            _fSurgeFl := fSlope * (fPress - fPressRef);                        (* 喘振流量下限 = 斜率 × (压力-参考)（乘性，无除零；可为负即无喘振约束） / Surge flow limit *)
            _fMargI := (fFlow - _fSurgeFl) / fFlowSpan;                        (* 归一化裕度：除子量程已过闸 [-] / Normalised margin *)
            IF _fMargI > DL_PSG_PCTMAX THEN
                _fMargI := DL_PSG_PCTMAX;                                      (* 裕度上限饱和 1（最后一次写） / Margin upper saturation *)
            ELSIF _fMargI < DL_PSG_PCTMIN THEN
                _fMargI := DL_PSG_PCTMIN;                                      (* 裕度下限饱和 0（最后一次写） / Margin lower saturation *)
            END_IF
            fMargin := _fMargI;                                                (* 裕度出口 / Margin outlet *)
            IF _fMargI < fMarginMin THEN
                bSurgeWarn := TRUE;                                            (* 裕度低于门槛：逼近告警（电平） / Margin below threshold *)
                _eCause := E_DL_PsgCause.eSurge;                               (* 成因更新：喘振逼近（诊断归因，非锁存故障） / Cause: surge proximity *)
                _fTarget := DL_PSG_DERMAX;                                     (* 降载目标 = 系数下限（深降载） / Target = derating floor *)
            ELSE
                _fTarget := DL_PSG_PCTMAX;                                     (* 裕度充足：恢复目标 = 全流量 / Target = full flow *)
            END_IF
            _fStep := fRampRate * _fDtSec;                                     (* 本拍斜坡步长（周期已过闸，REAL×REAL） / Ramp step *)
            IF _fFac < _fTarget THEN
                _fFac := _fFac + _fStep;                                       (* 恢复方向斜坡递增 / Ramp up *)
                IF _fFac > _fTarget THEN
                    _fFac := _fTarget;                                         (* 步长越目标即钳到目标（最后一次写） / Clamp to target *)
                END_IF
            ELSIF _fFac > _fTarget THEN
                _fFac := _fFac - _fStep;                                       (* 降载方向斜坡递减 / Ramp down *)
                IF _fFac < _fTarget THEN
                    _fFac := _fTarget;                                         (* 步长越目标即钳到目标（最后一次写） / Clamp to target *)
                END_IF
                IF _fFac < DL_PSG_DERMAX THEN
                    _fFac := DL_PSG_DERMAX;                                    (* 系数下限钳位（最后一次写） / Derating floor clamp *)
                END_IF
            END_IF
            fDerateFac := _fFac;                                               (* 系数出口（斜坡状态镜像） / Factor outlet *)
            IF ABS(fFlowCmd) > DL_PSG_EPS THEN                                 (* 流量命令有效才算限幅（除零前置，边界②） / Limit only with valid command *)
                fFlowLimit := fFlowCmd * _fFac;                                (* 限幅 = 命令 × 系数 [m3/h] / Limit = command times factor *)
            ELSE
                fFlowLimit := 0.0;                                             (* 命令近零：限幅 0（已充分降载语义） / Zero command: limit zero *)
            END_IF
        END_IF                                                                 (* 非有限输入：斜坡保持上拍值（边界③） / Non-finite: hold ramp *)
    E_DL_PsgState.eFault:                                                      (* 故障相：冻结保持末值，仅复位沿出 / Fault *)
        ;                                                                      (* 锁存回放（R28） / Replay from latch *)
    ELSE                                                                       (* 非法相位兜底迁安全态 / Illegal phase fallback *)
        _eState := E_DL_PsgState.eFault;                                       (* 迁故障相 / To fault *)
        _bFault := TRUE;                                                       (* 同步锁存 / Latch *)
        _eCause := E_DL_PsgCause.ePhaseBad;                                    (* 成因：非法相位 / Cause: illegal phase *)
END_CASE

(* —— 段 5：出口映射（bError/eState 同源，R191） —— *)
bError := _bFault;                                                             (* 故障标志镜像 / Fault flag mirror *)
eState := _eState;                                                             (* 状态出口 / State outlet *)
eCause := _eCause;                                                             (* 成因出口 / Cause outlet *)
END_FUNCTION_BLOCK

(* ---- FB_DL_PwmDutyController.st ---- *)
(*==============================================================================
 * 组件名称 (Component)  : FB_DL_PwmDutyController
 * 所属子库 (Sublibrary) : DL_Algo
 * 当前版本 (Version)    : 1.0.1
 * 兼容性   (Platform)   : CODESYS 3.5 / TwinCAT 3 / 汇川 InoProShop / Machine Expert
 *                         仅依赖 Standard.library（MIN / MAX / ABS），零厂商方言
 * 功能描述 (Function)   : 时间比例慢速 PWM 控制器。把 0~100% 占空比调制成周期级
 *                         布尔输出，驱动固态继电器（SSR）/接触器做加热功率调节，
 *                         避免高频开关对触点与电网的冲击。周期 tPeriod 内按占空比
 *                         分配导通时间；含最短导通/关断时间抑制（过窄脉冲跨周期
 *                         累加补偿，不足差额记入债务下周期叠加）、反相输出。
 *                         输出可与 PID 输出直连（0~100% 占空比）。
 * 开源溯源 (Origin)     : 原创实现。欠脉冲跨周期补偿思想源自 PID_Compact 的
 *                         脉冲发生器公开行为定义，clean-room 编写，
 *                         未复制任何厂商私有库源码。
 * 本文件内含       : TYPE  E_DL_PwmState（配套枚举，归属 DL_Algo）
 *                    FB    FB_DL_PwmDutyController
 * 依赖     (Depends)    : 无 DL_ 内部依赖；Standard.library: MIN / MAX / ABS
 * 红线自检 (Redline)    : R1 ✓ 零全局变量表与外部变量引用 ｜ R2 ✓ 零物理 IO 地址直写
 *                         R3 ✓ 纯 IEC 61131-3 ｜ R4 ✓ 周期/占空比/债务钳位
 *                         R5 ✓ 全变量中英双语同行注释 ｜ R6 ✓ 四态 ENUM+CASE+ELSE
 *                         R7 N/A（无定时器/边沿实例，相位自累加）
 * 【边界披露 / Boundary disclosure】
 *   B1 tPeriod < tMinOn + tMinOff：钳位 tPeriod := tMinOn + tMinOff 置 16#0002_0801。
 *   B2 tPeriod 低于 1s 下限：钳位到 1s 并置 16#0002_0801。
 *   B3 占空比越界钳位 0..100 置 16#0002_0001。
 *   B4 债务钳位 0..1 防无限累积；100% 占空比清空债务（全开无需补偿）。
 *   B5 使能跌落立即输出 FALSE 且债务清零，恢复后从周期起点重新计相位。
 *   B6 最短导通抑制：有效 ON 时间 < tMinOn 的窄脉冲并入债务，输出保持关断；
 *      最短关断抑制：OFF 间隙 < tMinOff 时合并为全周期导通（债务清零）。
 * 【验收向量 / Acceptance vectors】
 *   V1  fDuty=50，tPeriod=10S，tSampleTime=100MS → 每周期导通 5.0s、关断 5.0s，
 *       bPwmOut 方波占空比 50%，nCycleCount 每秒递增 0.1
 *   V2  fDuty=100 → bPwmOut 恒 TRUE、fDebt=0；fDuty=0 → 恒 FALSE
 *   V3  fDuty=0.2（ON 期望 20ms < tMinOn=500MS）→ 窄脉冲并入债务，bPwmOut 保持
 *       FALSE；连续 50 周期后债务足额释放为一个 ≥500ms 的长脉冲
 *   V4  fDuty=99.9（OFF 期望 10ms < tMinOff=500MS）→ 合并为全周期导通
 *   V5  tMinOn+tMinOff=12S > tPeriod=10S → tPeriod 钳位 12S、16#0002_0801
 *   V6  fDuty=150 → 钳位 100、16#0002_0001
 *   V7  bInvert=TRUE → bPwmOut 反相；bEnable=FALSE → bPwmOut 强制 FALSE
 * 修订历史 (Revision)   :
 *   2026-11-15  v1.0.0  首版入库（Round 04 · Phase 3 · DL_Algo 批次）
 *   2026-11-15  v1.0.1  阶段五终审精修：首次使能当拍立即结算占空比配额，
 *                       消除首周期无条件关断；bInit 由死变量转为有效标志
 *============================================================================*)

(*-----------------------------------------------------------------------------
 * 枚举: E_DL_PwmState（归属 DL_Algo，与 FB_DL_PwmDutyController 同文件）
 * 含义: 慢速 PWM 相位状态机。数值步长留空位便于后续插态而不破坏已有工程。
 *----------------------------------------------------------------------------*)
TYPE E_DL_PwmState :
(
    eIdle     := 0,   // 空闲态：未使能，输出关断 / Idle state, output off
    eOnPhase  := 10,  // 导通段：周期相位在有效占空比区间内 / On phase, cycle phase within effective duty
    eOffPhase := 20,  // 关断段：周期相位超出有效占空比区间 / Off phase, phase beyond effective duty
    eFault    := 99   // 故障兜底态：非法状态拦截，自动回空闲 / Fault fallback, auto recover to idle
);
END_TYPE

(*==============================================================================
 * 功能块: FB_DL_PwmDutyController
 * 调用约定: 每个扫描周期无条件调用一次；占空比可在周期中途修改，下周期生效配额。
 * 无状态泄漏: 全部状态驻留于实例私有 VAR，可多实例并行互不影响。
 * 相位披露: fPhase 每拍累加 fDt/fPeriod，达到 1.0 回卷并结算本周期配额；
 *           输出与 PID 占空比直连，脉宽分辨率 = 扫描周期（慢速 PWM 语义）。
 *============================================================================*)
FUNCTION_BLOCK FB_DL_PwmDutyController
VAR_INPUT
    bEnable     : BOOL := FALSE;      // 使能标志，FALSE 立即关断并清债务 / Enable flag, FALSE forces off and clears debt
    fDuty       : REAL := 0.0;        // 占空比输入 [%]，0..100，越界钳位 / Duty cycle input [%], 0..100 clamped
    tPeriod     : TIME := T#10S;      // PWM 周期 [s]，下限 1s 且须 >= 最短开关时间和 / PWM period [s], min 1s
    tMinOn      : TIME := T#500MS;    // 最短导通时间 [s]，窄脉冲并入债务 / Minimum on time [s], narrow pulses deferred
    tMinOff     : TIME := T#500MS;    // 最短关断时间 [s]，两者之和须 < tPeriod / Minimum off time [s]
    bInvert     : BOOL := FALSE;      // 反相输出，TRUE 时输出取反 / Invert output, TRUE inverts the boolean
    tSampleTime : TIME := T#100MS;    // 采样周期 [s]，小于 10ms 钳位为 10ms / Sample time [s], clamped to 10ms
END_VAR
VAR_OUTPUT
    bPwmOut     : BOOL;               // PWM 布尔输出（已含反相处理） / PWM boolean output, invert applied
    fDutyEff    : REAL;               // 本周期实际有效占空比 [%]，含债务补偿 / Effective duty this cycle [%] with debt
    nCycleCount : UDINT;              // 已完成周期计数 [个] / Completed cycle count
    bError      : BOOL;               // 故障标志（瞬时，逐拍重算） / Fault flag, transient, recomputed every scan
    uErrorId    : UDINT;              // 故障码，0 = 无故障 / Error code, 0 = no error
END_VAR
VAR
    fPhase      : REAL;               // 周期相位 [0..1] / Cycle phase [0..1]
    fDutyEffInt : REAL;               // 本周期有效占空比（内部小数）[0..1] / Effective duty fraction [0..1]
    fDebt       : REAL;               // 欠脉冲债务 [0..1]，跨周期累加 / Pulse debt [0..1], accumulated across cycles
    bOnState    : BOOL;               // 原始导通状态（未反相） / Raw on state before inversion
    fPeriodSec  : REAL;               // 钳位后周期 [s] / Clamped period [s]
    fMinOnSec   : REAL;               // 最短导通时间 [s] / Minimum on time [s]
    fMinOffSec  : REAL;               // 最短关断时间 [s] / Minimum off time [s]
    fDt         : REAL;               // 折算后的采样周期 [s] / Converted sample period [s]
    fDutyC      : REAL;               // 钳位后占空比 [%] / Clamped duty [%]
    fDutyReq    : REAL;               // 本周期占空比请求（含债务）[0..1] / Duty request with debt [0..1]
    tPeriodEff  : TIME;               // 钳位后周期时刻值 / Clamped period time value
    bInit       : BOOL;               // 首扫标志，FALSE 触发配额立即结算 / First-scan flag, FALSE settles quota immediately
    eState      : E_DL_PwmState;      // 主状态机当前状态 / Current state of the main state machine
END_VAR
VAR CONSTANT
    DL_PWM_DUTY_MAX   : REAL := 100.0;  // 占空比上限 [%] / Duty cycle upper limit [%]
    DL_PWM_PERIOD_MIN : TIME := T#1S;   // 周期下限 [s] / Period lower limit [s]
END_VAR

(*------------------------------------------------------------------------------
 * 段 1｜公共参数处理（通用约定 0-1）：周期钳位、故障码瞬时清零
 *      Common handling: period clamp, transient error code reset
 *-----------------------------------------------------------------------------*)
uErrorId := 16#0000_0000;               // 故障码逐拍重算 / Error code recomputed every scan
bError   := FALSE;                      // 故障标志逐拍重算 / Fault flag recomputed every scan

IF tSampleTime < T#10MS THEN
    fDt      := TIME_TO_REAL(T#10MS) / 1000.0; // 非法周期钳位为 10ms / Illegal period clamped to 10ms
    uErrorId := 16#0002_0002;           // 采样周期非法已钳位 / Sample time illegal, clamped
ELSE
    fDt      := TIME_TO_REAL(tSampleTime) / 1000.0; // 周期换算为秒 [s] / Period converted to seconds [s]
END_IF

(*------------------------------------------------------------------------------
 * 段 2｜周期钳位（边界 B1/B2）：先保证 >= 最短开关时间和，再保证 >= 1s 下限
 *      Period clamping: ensure >= min on+off sum first, then >= 1s floor
 *-----------------------------------------------------------------------------*)
tPeriodEff := tPeriod;                  // 周期初值 / Initial period value
IF tMinOn + tMinOff > tPeriodEff THEN
    tPeriodEff := tMinOn + tMinOff;     // 周期放大到最短开关时间和 / Period raised to min on+off sum
    uErrorId   := 16#0002_0801;         // 周期小于最短开关时间和已钳位 / Period below min on+off sum, clamped
END_IF
IF tPeriodEff < DL_PWM_PERIOD_MIN THEN
    tPeriodEff := DL_PWM_PERIOD_MIN;    // 周期放大到 1s 下限 / Period raised to 1s floor
    uErrorId   := 16#0002_0801;         // 周期非法已钳位 / Period illegal, clamped
END_IF

fPeriodSec := TIME_TO_REAL(tPeriodEff) / 1000.0; // 周期换算为秒 [s] / Period converted to seconds [s]
fMinOnSec  := TIME_TO_REAL(tMinOn) / 1000.0;     // 最短导通换算为秒 [s] / Min on time in seconds [s]
fMinOffSec := TIME_TO_REAL(tMinOff) / 1000.0;    // 最短关断换算为秒 [s] / Min off time in seconds [s]

(*------------------------------------------------------------------------------
 * 段 3｜占空比钳位（边界 B3）：0..100，越界告警不中断
 *      Duty clamping: 0..100, over-range warns without stopping
 *-----------------------------------------------------------------------------*)
fDutyC := fDuty;                        // 占空比初值 / Initial duty value
IF fDutyC < 0.0 THEN
    fDutyC   := 0.0;                    // 下越界钳位 / Under-range clamped
    uErrorId := 16#0002_0001;           // 参数越界已钳位 / Parameter out of range, clamped
END_IF
IF fDutyC > DL_PWM_DUTY_MAX THEN
    fDutyC   := DL_PWM_DUTY_MAX;        // 上越界钳位 / Over-range clamped
    uErrorId := 16#0002_0001;           // 参数越界已钳位 / Parameter out of range, clamped
END_IF

(*------------------------------------------------------------------------------
 * 段 4｜使能失效语义（边界 B5）：立即关断、清债务、相位归零、回空闲
 *      Disabled semantics: immediate off, debt cleared, phase reset, idle
 *-----------------------------------------------------------------------------*)
IF NOT bEnable THEN
    bPwmOut     := FALSE;               // 输出强制关断（反相不生效，安全优先）/ Output forced off, invert bypassed for safety
    bOnState    := FALSE;               // 原始导通状态清零 / Raw on state cleared
    fPhase      := 0.0;                 // 相位归零 / Phase reset
    fDebt       := 0.0;                 // 债务清零 / Debt cleared
    fDutyEffInt := 0.0;                 // 本周期有效占空比清零 / Effective duty cleared
    fDutyEff    := 0.0;                 // 输出占空比清零 / Output duty cleared
    eState      := eIdle;               // 强制空闲 / Force idle
    bInit       := FALSE;               // 复位首扫标志，重使能当拍立即结算配额 / Reset init flag, settle quota on re-enable
ELSE
    (*--------------------------------------------------------------------------
     * 段 5a｜相位推进与周期结算：fPhase >= 1.0 回卷，结算本周期配额
     *     Phase advance and cycle settlement: wrap at 1.0, settle quota
     *-------------------------------------------------------------------------*)
    fPhase := fPhase + fDt / fPeriodSec; // 相位累加 [0..1] / Phase accumulation [0..1]

    IF (fPhase >= 1.0) OR (NOT bInit) THEN
        IF fPhase >= 1.0 THEN
            fPhase := fPhase - 1.0;     // 相位回卷 / Phase wrapped
            IF fPhase >= 1.0 THEN
                fPhase := 0.0;          // 单拍跨度超周期时强制归零（防御）/ Forced reset if one scan exceeds period
            END_IF
        END_IF

        fDutyReq := fDutyC / DL_PWM_DUTY_MAX + fDebt; // 占空比请求含债务 [0..1] / Duty request with debt [0..1]
        fDutyEffInt := MIN(fDutyReq, 1.0);            // 本周期配额上限 100% / Cycle quota capped at 100%
        fDebt := fDutyReq - fDutyEffInt;              // 剩余债务 / Remaining debt
        fDebt := MIN(MAX(fDebt, 0.0), 1.0);           // 债务钳位防无限累积 / Debt clamped against runaway

        (* 最短导通抑制（边界 B6 前半）：窄脉冲并入债务 / Min-on suppression: narrow pulse merged into debt *)
        IF (fDutyEffInt > 0.0) AND (fDutyEffInt * fPeriodSec < fMinOnSec) THEN
            fDebt       := MIN(fDebt + fDutyEffInt, 1.0); // 窄脉冲差额记账 / Narrow pulse booked into debt
            fDutyEffInt := 0.0;                            // 本周期保持关断 / Cycle held off
        END_IF

        (* 最短关断抑制（边界 B6 后半）：OFF 间隙过窄合并为全开 / Min-off suppression: narrow gap merged to full on *)
        IF (fDutyEffInt < 1.0) AND ((1.0 - fDutyEffInt) * fPeriodSec < fMinOffSec) THEN
            fDutyEffInt := 1.0;         // 合并为全周期导通 / Merged to full-cycle on
            fDebt       := 0.0;         // 全开无需补偿，债务清零 / Debt cleared, full on needs no compensation
        END_IF

        fDutyEff := fDutyEffInt * DL_PWM_DUTY_MAX; // 有效占空比输出 [%] / Effective duty output [%]
        nCycleCount := nCycleCount + 1;             // 周期计数递增 / Cycle count incremented
        bInit := TRUE;                              // 首扫配额已结算 / Initial quota settled
    END_IF

    (*--------------------------------------------------------------------------
     * 段 5b｜主状态机（红线 R6）：四态 ENUM + CASE + ELSE 兜底，相位派生覆盖
     *     Main state machine: four-state ENUM + CASE with phase-derived coverage
     *-------------------------------------------------------------------------*)
    CASE eState OF

        eIdle:  // 空闲态：使能后按相位派生进入导通或关断段 / Idle: derive on/off phase after enable
            IF fPhase < fDutyEffInt THEN
                eState := eOnPhase;     // 相位在配额内，导通 / Phase within quota, on
            ELSE
                eState := eOffPhase;    // 相位超配额，关断 / Phase beyond quota, off
            END_IF

        eOnPhase:  // 导通段：相位越过配额即切换关断 / On phase: switch off when phase exceeds quota
            IF fPhase >= fDutyEffInt THEN
                eState := eOffPhase;    // 切换到关断段 / Switch to off phase
            END_IF

        eOffPhase:  // 关断段：新周期配额生效即切换导通 / Off phase: switch on when new quota applies
            IF fPhase < fDutyEffInt THEN
                eState := eOnPhase;     // 切换到导通段 / Switch to on phase
            END_IF

        eFault:  // 故障兜底态：无复位引脚，当拍回空闲重派生 / Fault fallback: recover to idle, re-derive
            eState := eIdle;            // 自动恢复空闲 / Auto recover to idle

        ELSE  // 非法状态拦截：任何未定义状态一律进故障态并置码 / Illegal state interception
            eState   := eFault;         // 强制故障态 / Force fault state
            uErrorId := 16#0002_0005;   // 非法状态兜底 / Illegal state fallback
            bError   := TRUE;           // 故障标志置位 / Fault flag set

    END_CASE;

    bOnState := (eState = eOnPhase);    // 原始导通状态派生 / Raw on state derived
    bPwmOut  := (bOnState <> bInvert);  // 反相处理后输出 / Output after inversion
END_IF
END_FUNCTION_BLOCK
